Universal Robots URScript: FaiChun_9 Jan_11_2_t2.script

def Machining1():
  # Default parameters:
  global speed_ms = 0.05
  global speed_rads = 0.75
  global accel_mss = 3
  global accel_radss = 1.2
  global blend_radius_m = 0.0003

  # Add subprograms here
  # Start of main program
  # Program generated by RoboDK v5.6.8 for UR10e on 17/01/2025 16:04:48
  # Using nominal kinematics.
  blend_radius_m = 0.0003
  speed_ms = 0.05
  # set_reference(p[0.340000, -0.053000, 0.001500, 0.000000, 0.000000, 0.000000])
  set_tcp(p[0.000000, 0.000000, 0.252000, 0.000000, 0.000000, 0.000000])
  # Show Tool
  movej([0.537356, -1.385611, -2.455322, -0.871456, 1.570796, 2.108152],accel_radss,speed_rads,0,blend_radius_m)
  movel([0.537356, -1.438776, -2.485556, -0.788057, 1.570796, 2.108152],accel_mss,speed_ms,0,blend_radius_m)
  #SetTool1
  #M_RunCode6
  #SetRPM60000
  speed_ms = 0.05
  #M_RunCode3
  movel([0.537356, -1.461982, -2.496787, -0.753620, 1.570796, 2.108152],accel_mss,speed_ms,0,blend_radius_m)
  speed_ms = 0.003
  movel([0.537356, -1.467978, -2.499523, -0.744888, 1.570796, 2.108152],accel_mss,speed_ms,0,blend_radius_m)
  speed_ms = 0.02
  movel([0.264301, -1.461173, -2.505187, -0.746029, 1.570796, 1.835098],accel_mss,speed_ms,0,blend_radius_m)
  movel([0.376012, -1.125586, -2.705707, -0.881096, 1.570796, 1.946808],accel_mss,speed_ms,0,blend_radius_m)
  movel([0.747752, -1.141566, -2.699168, -0.871655, 1.570796, 2.318548],accel_mss,speed_ms,0,blend_radius_m)
  movel([0.537356, -1.467978, -2.499523, -0.744888, 1.570796, 2.108152],accel_mss,speed_ms,0,blend_radius_m)
  speed_ms = 0.003
  movel([0.537356, -1.461982, -2.496787, -0.753620, 1.570796, 2.108152],accel_mss,speed_ms,0,blend_radius_m)
  speed_ms = 0.05
  movel([0.537356, -1.438776, -2.485556, -0.788057, 1.570796, 2.108152],accel_mss,speed_ms,0,blend_radius_m)
  #M_RunCode9
  movel([0.537227, -1.429917, -2.492594, -0.789878, 1.570796, 2.108023],accel_mss,speed_ms,0,blend_radius_m)
  #M_RunCode3
  movel([0.537227, -1.453304, -2.503930, -0.755154, 1.570796, 2.108023],accel_mss,speed_ms,0,blend_radius_m)
  speed_ms = 0.003
  movel([0.537227, -1.459350, -2.506693, -0.746346, 1.570796, 2.108023],accel_mss,speed_ms,0,blend_radius_m)
  speed_ms = 0.012
  movel([0.533373, -1.458727, -2.507206, -0.746456, 1.570796, 2.104169],accel_mss,speed_ms,0,blend_radius_m)
  movel([0.531104, -1.462629, -2.503981, -0.745779, 1.570796, 2.101900],accel_mss,speed_ms,0,blend_radius_m)
  movel([0.525395, -1.461744, -2.504715, -0.745930, 1.570796, 2.096191],accel_mss,speed_ms,0,blend_radius_m)
  movel([0.527644, -1.457831, -2.507943, -0.746615, 1.570796, 2.098440],accel_mss,speed_ms,0,blend_radius_m)
  movel([0.525630, -1.457526, -2.508194, -0.746669, 1.570796, 2.096426],accel_mss,speed_ms,0,blend_radius_m)
  movel([0.523386, -1.461442, -2.504965, -0.745982, 1.570796, 2.094182],accel_mss,speed_ms,0,blend_radius_m)
  movel([0.518575, -1.460738, -2.505547, -0.746104, 1.570796, 2.089372],accel_mss,speed_ms,0,blend_radius_m)
  movel([0.517641, -1.460602, -2.505659, -0.746128, 1.570796, 2.088438],accel_mss,speed_ms,0,blend_radius_m)
  movel([0.520940, -1.454785, -2.510440, -0.747164, 1.570796, 2.091736],accel_mss,speed_ms,0,blend_radius_m)
  movel([0.524842, -1.455357, -2.509972, -0.747060, 1.570796, 2.095639],accel_mss,speed_ms,0,blend_radius_m)
  movel([0.526016, -1.453307, -2.511646, -0.747436, 1.570796, 2.096813],accel_mss,speed_ms,0,blend_radius_m)
  movel([0.520074, -1.452441, -2.512352, -0.747596, 1.570796, 2.090870],accel_mss,speed_ms,0,blend_radius_m)
  movel([0.515622, -1.460318, -2.505894, -0.746177, 1.570796, 2.086418],accel_mss,speed_ms,0,blend_radius_m)
  movel([0.514683, -1.460189, -2.506001, -0.746199, 1.570796, 2.085480],accel_mss,speed_ms,0,blend_radius_m)
  speed_ms = 0.02
  movel([0.406474, -1.451431, -2.513173, -0.747785, 1.570796, 1.977270],accel_mss,speed_ms,0,blend_radius_m)
  movel([0.291548, -1.454758, -2.510462, -0.747169, 1.570796, 1.862344],accel_mss,speed_ms,0,blend_radius_m)
  speed_ms = 0.012
  movel([0.294155, -1.446765, -2.516946, -0.748678, 1.570796, 1.864951],accel_mss,speed_ms,0,blend_radius_m)
  movel([0.287539, -1.447324, -2.516496, -0.748569, 1.570796, 1.858335],accel_mss,speed_ms,0,blend_radius_m)
  movel([0.286869, -1.449403, -2.514817, -0.748169, 1.570796, 1.857666],accel_mss,speed_ms,0,blend_radius_m)
  movel([0.291218, -1.449032, -2.515117, -0.748240, 1.570796, 1.862014],accel_mss,speed_ms,0,blend_radius_m)
  movel([0.289302, -1.454935, -2.510317, -0.747137, 1.570796, 1.860098],accel_mss,speed_ms,0,blend_radius_m)
  movel([0.288263, -1.455022, -2.510246, -0.747121, 1.570796, 1.859059],accel_mss,speed_ms,0,blend_radius_m)
  movel([0.282904, -1.455482, -2.509870, -0.747037, 1.570796, 1.853700],accel_mss,speed_ms,0,blend_radius_m)
  movel([0.284166, -1.451508, -2.513110, -0.747771, 1.570796, 1.854962],accel_mss,speed_ms,0,blend_radius_m)
  movel([0.281913, -1.451708, -2.512947, -0.747733, 1.570796, 1.852710],accel_mss,speed_ms,0,blend_radius_m)
  movel([0.280661, -1.455682, -2.509706, -0.747001, 1.570796, 1.851457],accel_mss,speed_ms,0,blend_radius_m)
  movel([0.274256, -1.456275, -2.509221, -0.746894, 1.570796, 1.845052],accel_mss,speed_ms,0,blend_radius_m)
  movel([0.275479, -1.452309, -2.512459, -0.747621, 1.570796, 1.846276],accel_mss,speed_ms,0,blend_radius_m)
  movel([0.271129, -1.452735, -2.512112, -0.747542, 1.570796, 1.841925],accel_mss,speed_ms,0,blend_radius_m)
  movel([0.272932, -1.446825, -2.516897, -0.748666, 1.570796, 1.843728],accel_mss,speed_ms,0,blend_radius_m)
  movel([0.277309, -1.446393, -2.517245, -0.748750, 1.570796, 1.848106],accel_mss,speed_ms,0,blend_radius_m)
  movel([0.277957, -1.444307, -2.518920, -0.749161, 1.570796, 1.848754],accel_mss,speed_ms,0,blend_radius_m)
  movel([0.273570, -1.444740, -2.518573, -0.749076, 1.570796, 1.844366],accel_mss,speed_ms,0,blend_radius_m)
  movel([0.275104, -1.439738, -2.522566, -0.750085, 1.570796, 1.845900],accel_mss,speed_ms,0,blend_radius_m)
  movel([0.275407, -1.438760, -2.523343, -0.750287, 1.570796, 1.846203],accel_mss,speed_ms,0,blend_radius_m)
  movel([0.281948, -1.438112, -2.523856, -0.750421, 1.570796, 1.852744],accel_mss,speed_ms,0,blend_radius_m)
  movel([0.280675, -1.442163, -2.520635, -0.749591, 1.570796, 1.851471],accel_mss,speed_ms,0,blend_radius_m)
  movel([0.282958, -1.441947, -2.520808, -0.749635, 1.570796, 1.853754],accel_mss,speed_ms,0,blend_radius_m)
  movel([0.284909, -1.435781, -2.525698, -0.750910, 1.570796, 1.855706],accel_mss,speed_ms,0,blend_radius_m)
  movel([0.276057, -1.436649, -2.525013, -0.750727, 1.570796, 1.846853],accel_mss,speed_ms,0,blend_radius_m)
  movel([0.315010, -1.315779, -2.609859, -0.786751, 1.570796, 1.885806],accel_mss,speed_ms,0,blend_radius_m)
  speed_ms = 0.02
  movel([0.366945, -1.166741, -2.688352, -0.857296, 1.570796, 1.937742],accel_mss,speed_ms,0,blend_radius_m)
  movel([0.367496, -1.165223, -2.689023, -0.858143, 1.570796, 1.938292],accel_mss,speed_ms,0,blend_radius_m)
  speed_ms = 0.012
  movel([0.379333, -1.163455, -2.689801, -0.859133, 1.570796, 1.950130],accel_mss,speed_ms,0,blend_radius_m)
  movel([0.382947, -1.153742, -2.694017, -0.864630, 1.570796, 1.953743],accel_mss,speed_ms,0,blend_radius_m)
  movel([0.379852, -1.154196, -2.693822, -0.864371, 1.570796, 1.950648],accel_mss,speed_ms,0,blend_radius_m)
  movel([0.377482, -1.160600, -2.691050, -0.860739, 1.570796, 1.948278],accel_mss,speed_ms,0,blend_radius_m)
  movel([0.368695, -1.161928, -2.690470, -0.859991, 1.570796, 1.939492],accel_mss,speed_ms,0,blend_radius_m)
  movel([0.369247, -1.160401, -2.691137, -0.860851, 1.570796, 1.940044],accel_mss,speed_ms,0,blend_radius_m)
  movel([0.372128, -1.152454, -2.694569, -0.865366, 1.570796, 1.942924],accel_mss,speed_ms,0,blend_radius_m)
  movel([0.378119, -1.151528, -2.694965, -0.865896, 1.570796, 1.948915],accel_mss,speed_ms,0,blend_radius_m)
  movel([0.379358, -1.148166, -2.696395, -0.867829, 1.570796, 1.950154],accel_mss,speed_ms,0,blend_radius_m)
  movel([0.373347, -1.149100, -2.695999, -0.867291, 1.570796, 1.944143],accel_mss,speed_ms,0,blend_radius_m)
  movel([0.376872, -1.139423, -2.700060, -0.872907, 1.570796, 1.947669],accel_mss,speed_ms,0,blend_radius_m)
  movel([0.382941, -1.138466, -2.700456, -0.873467, 1.570796, 1.953738],accel_mss,speed_ms,0,blend_radius_m)
  movel([0.385401, -1.131831, -2.703181, -0.877377, 1.570796, 1.956197],accel_mss,speed_ms,0,blend_radius_m)
  movel([0.394435, -1.130456, -2.703741, -0.878193, 1.570796, 1.965231],accel_mss,speed_ms,0,blend_radius_m)
  movel([0.391917, -1.137114, -2.701015, -0.874260, 1.570796, 1.962713],accel_mss,speed_ms,0,blend_radius_m)
  movel([0.395057, -1.136658, -2.701203, -0.874528, 1.570796, 1.965853],accel_mss,speed_ms,0,blend_radius_m)
  movel([0.397596, -1.129993, -2.703928, -0.878468, 1.570796, 1.968392],accel_mss,speed_ms,0,blend_radius_m)
  movel([0.406602, -1.128726, -2.704442, -0.879221, 1.570796, 1.977398],accel_mss,speed_ms,0,blend_radius_m)
  movel([0.402769, -1.138603, -2.700399, -0.873387, 1.570796, 1.973565],accel_mss,speed_ms,0,blend_radius_m)
  movel([0.396746, -1.139429, -2.700057, -0.872903, 1.570796, 1.967543],accel_mss,speed_ms,0,blend_radius_m)
  movel([0.395440, -1.142849, -2.698632, -0.870908, 1.570796, 1.966236],accel_mss,speed_ms,0,blend_radius_m)
  movel([0.404555, -1.141619, -2.699146, -0.871624, 1.570796, 1.975351],accel_mss,speed_ms,0,blend_radius_m)
  movel([0.409752, -1.128301, -2.704613, -0.879474, 1.570796, 1.980548],accel_mss,speed_ms,0,blend_radius_m)
  movel([0.568735, -1.120522, -2.707727, -0.884139, 1.570796, 2.139531],accel_mss,speed_ms,0,blend_radius_m)
  speed_ms = 0.02
  movel([0.712082, -1.141087, -2.699368, -0.871934, 1.570796, 2.282879],accel_mss,speed_ms,0,blend_radius_m)
  movel([0.703666, -1.154003, -2.693905, -0.864481, 1.570796, 2.274462],accel_mss,speed_ms,0,blend_radius_m)
  speed_ms = 0.012
  movel([0.711078, -1.155876, -2.693099, -0.863414, 1.570796, 2.281874],accel_mss,speed_ms,0,blend_radius_m)
  movel([0.713256, -1.152569, -2.694520, -0.865300, 1.570796, 2.284052],accel_mss,speed_ms,0,blend_radius_m)
  movel([0.708376, -1.151318, -2.695054, -0.866017, 1.570796, 2.279173],accel_mss,speed_ms,0,blend_radius_m)
  movel([0.714644, -1.141751, -2.699091, -0.871547, 1.570796, 2.285440],accel_mss,speed_ms,0,blend_radius_m)
  movel([0.715827, -1.142057, -2.698963, -0.871369, 1.570796, 2.286624],accel_mss,speed_ms,0,blend_radius_m)
  movel([0.721900, -1.143661, -2.698292, -0.870436, 1.570796, 2.292696],accel_mss,speed_ms,0,blend_radius_m)
  movel([0.717633, -1.150105, -2.695571, -0.866713, 1.570796, 2.288429],accel_mss,speed_ms,0,blend_radius_m)
  movel([0.720150, -1.150783, -2.695282, -0.866323, 1.570796, 2.290946],accel_mss,speed_ms,0,blend_radius_m)
  movel([0.724433, -1.144348, -2.698004, -0.870037, 1.570796, 2.295229],accel_mss,speed_ms,0,blend_radius_m)
  movel([0.731605, -1.146355, -2.697160, -0.868874, 1.570796, 2.302401],accel_mss,speed_ms,0,blend_radius_m)
  movel([0.727300, -1.152759, -2.694438, -0.865192, 1.570796, 2.298096],accel_mss,speed_ms,0,blend_radius_m)
  movel([0.732091, -1.154132, -2.693850, -0.864408, 1.570796, 2.302888],accel_mss,speed_ms,0,blend_radius_m)
  movel([0.725789, -1.163458, -2.689799, -0.859132, 1.570796, 2.296585],accel_mss,speed_ms,0,blend_radius_m)
  movel([0.721022, -1.162117, -2.690387, -0.859885, 1.570796, 2.291818],accel_mss,speed_ms,0,blend_radius_m)
  movel([0.718847, -1.165363, -2.688961, -0.858065, 1.570796, 2.289644],accel_mss,speed_ms,0,blend_radius_m)
  movel([0.723604, -1.166697, -2.688372, -0.857320, 1.570796, 2.294400],accel_mss,speed_ms,0,blend_radius_m)
  movel([0.718442, -1.174360, -2.684951, -0.853078, 1.570796, 2.289239],accel_mss,speed_ms,0,blend_radius_m)
  movel([0.717449, -1.175836, -2.684285, -0.852268, 1.570796, 2.288246],accel_mss,speed_ms,0,blend_radius_m)
  movel([0.710428, -1.173922, -2.685148, -0.853319, 1.570796, 2.281224],accel_mss,speed_ms,0,blend_radius_m)
  movel([0.714548, -1.167736, -2.687912, -0.856742, 1.570796, 2.285344],accel_mss,speed_ms,0,blend_radius_m)
  movel([0.712062, -1.167070, -2.688207, -0.857112, 1.570796, 2.282858],accel_mss,speed_ms,0,blend_radius_m)
  movel([0.705834, -1.176462, -2.684002, -0.851925, 1.570796, 2.276630],accel_mss,speed_ms,0,blend_radius_m)
  movel([0.715315, -1.179011, -2.682845, -0.850533, 1.570796, 2.286112],accel_mss,speed_ms,0,blend_radius_m)
  speed_ms = 0.02
  movel([0.619516, -1.325160, -2.604003, -0.783226, 1.570796, 2.190312],accel_mss,speed_ms,0,blend_radius_m)
  movel([0.546569, -1.443533, -2.519541, -0.749316, 1.570796, 2.117365],accel_mss,speed_ms,0,blend_radius_m)
  speed_ms = 0.012
  movel([0.538730, -1.442256, -2.520561, -0.749572, 1.570796, 2.109526],accel_mss,speed_ms,0,blend_radius_m)
  movel([0.535189, -1.448324, -2.515689, -0.748376, 1.570796, 2.105985],accel_mss,speed_ms,0,blend_radius_m)
  movel([0.537216, -1.448646, -2.515429, -0.748314, 1.570796, 2.108012],accel_mss,speed_ms,0,blend_radius_m)
  movel([0.539548, -1.444662, -2.518636, -0.749091, 1.570796, 2.110344],accel_mss,speed_ms,0,blend_radius_m)
  movel([0.545329, -1.445610, -2.517875, -0.748904, 1.570796, 2.116125],accel_mss,speed_ms,0,blend_radius_m)
  movel([0.544761, -1.446568, -2.517104, -0.748716, 1.570796, 2.115557],accel_mss,speed_ms,0,blend_radius_m)
  movel([0.541852, -1.451489, -2.513125, -0.747774, 1.570796, 2.112648],accel_mss,speed_ms,0,blend_radius_m)
  movel([0.537972, -1.450854, -2.513641, -0.747894, 1.570796, 2.108768],accel_mss,speed_ms,0,blend_radius_m)
  movel([0.536771, -1.452905, -2.511974, -0.747510, 1.570796, 2.107567],accel_mss,speed_ms,0,blend_radius_m)
  movel([0.540646, -1.453538, -2.511458, -0.747393, 1.570796, 2.111442],accel_mss,speed_ms,0,blend_radius_m)
  movel([0.537227, -1.459350, -2.506693, -0.746346, 1.570796, 2.108023],accel_mss,speed_ms,0,blend_radius_m)
  speed_ms = 0.003
  movel([0.537227, -1.453304, -2.503930, -0.755154, 1.570796, 2.108023],accel_mss,speed_ms,0,blend_radius_m)
  speed_ms = 0.05
  movel([0.537227, -1.429917, -2.492594, -0.789878, 1.570796, 2.108023],accel_mss,speed_ms,0,blend_radius_m)
  #M_RunCode9
  movel([0.423144, -1.170555, -2.652350, -0.889483, 1.570796, 1.993941],accel_mss,speed_ms,0,blend_radius_m)
  #M_RunCode3
  # num 0 inside
  movel([0.423144, -1.197858, -2.667024, -0.847507, 1.570796, 1.993941],accel_mss,speed_ms,0,blend_radius_m)
  speed_ms = 0.003
  movel([0.423144, -1.205044, -2.670628, -0.836717, 1.570796, 1.993941],accel_mss,speed_ms,0,blend_radius_m)
  speed_ms = 0.015
  movel([0.414451, -1.211707, -2.667382, -0.833300, 1.570796, 1.985247],accel_mss,speed_ms,0,blend_radius_m)
  movel([0.408145, -1.215978, -2.665275, -0.831136, 1.570796, 1.978941],accel_mss,speed_ms,0,blend_radius_m)
  movel([0.405824, -1.217205, -2.664666, -0.830518, 1.570796, 1.976621],accel_mss,speed_ms,0,blend_radius_m)
  movel([0.403998, -1.217788, -2.664376, -0.830225, 1.570796, 1.974795],accel_mss,speed_ms,0,blend_radius_m)
  movel([0.402664, -1.217733, -2.664403, -0.830253, 1.570796, 1.973460],accel_mss,speed_ms,0,blend_radius_m)
  movel([0.401818, -1.217039, -2.664748, -0.830602, 1.570796, 1.972614],accel_mss,speed_ms,0,blend_radius_m)
  movel([0.401559, -1.215868, -2.665329, -0.831191, 1.570796, 1.972356],accel_mss,speed_ms,0,blend_radius_m)
  movel([0.401991, -1.214387, -2.666062, -0.831940, 1.570796, 1.972787],accel_mss,speed_ms,0,blend_radius_m)
  movel([0.403116, -1.212593, -2.666947, -0.832850, 1.570796, 1.973912],accel_mss,speed_ms,0,blend_radius_m)
  movel([0.404937, -1.210479, -2.667984, -0.833926, 1.570796, 1.975733],accel_mss,speed_ms,0,blend_radius_m)
  movel([0.410670, -1.205076, -2.670613, -0.836701, 1.570796, 1.981466],accel_mss,speed_ms,0,blend_radius_m)
  movel([0.419217, -1.197936, -2.674037, -0.840416, 1.570796, 1.990013],accel_mss,speed_ms,0,blend_radius_m)
  movel([0.428065, -1.191105, -2.677261, -0.844024, 1.570796, 1.998861],accel_mss,speed_ms,0,blend_radius_m)
  movel([0.434586, -1.186692, -2.679317, -0.846381, 1.570796, 2.005382],accel_mss,speed_ms,0,blend_radius_m)
  movel([0.436993, -1.185433, -2.679899, -0.847057, 1.570796, 2.007789],accel_mss,speed_ms,0,blend_radius_m)
  movel([0.438876, -1.184846, -2.680170, -0.847373, 1.570796, 2.009672],accel_mss,speed_ms,0,blend_radius_m)
  movel([0.440232, -1.184936, -2.680129, -0.847325, 1.570796, 2.011028],accel_mss,speed_ms,0,blend_radius_m)
  movel([0.441059, -1.185700, -2.679775, -0.846913, 1.570796, 2.011856],accel_mss,speed_ms,0,blend_radius_m)
  movel([0.441266, -1.186954, -2.679195, -0.846240, 1.570796, 2.012062],accel_mss,speed_ms,0,blend_radius_m)
  movel([0.440764, -1.188513, -2.678471, -0.845406, 1.570796, 2.011560],accel_mss,speed_ms,0,blend_radius_m)
  movel([0.439549, -1.190375, -2.677602, -0.844412, 1.570796, 2.010346],accel_mss,speed_ms,0,blend_radius_m)
  movel([0.437636, -1.192534, -2.676590, -0.843265, 1.570796, 2.008432],accel_mss,speed_ms,0,blend_radius_m)
  movel([0.431736, -1.197976, -2.674018, -0.840395, 1.570796, 2.002532],accel_mss,speed_ms,0,blend_radius_m)
  movel([0.423144, -1.205044, -2.670628, -0.836717, 1.570796, 1.993941],accel_mss,speed_ms,0,blend_radius_m)
  speed_ms = 0.003
  movel([0.423144, -1.197858, -2.667024, -0.847507, 1.570796, 1.993941],accel_mss,speed_ms,0,blend_radius_m)
  speed_ms = 0.05
  movel([0.423144, -1.170555, -2.652350, -0.889483, 1.570796, 1.993941],accel_mss,speed_ms,0,blend_radius_m)
  #M_RunCode9
  movel([0.427307, -1.178294, -2.648743, -0.885352, 1.570796, 1.998103],accel_mss,speed_ms,0,blend_radius_m)
  #M_RunCode3
  #num 0 outside
  movel([0.427307, -1.205537, -2.663314, -0.843537, 1.570796, 1.998103],accel_mss,speed_ms,0,blend_radius_m)
  speed_ms = 0.003
  movel([0.427307, -1.212702, -2.666893, -0.832794, 1.570796, 1.998103],accel_mss,speed_ms,0,blend_radius_m)
  speed_ms = 0.015
  movel([0.424140, -1.215057, -2.665731, -0.831601, 1.570796, 1.994936],accel_mss,speed_ms,0,blend_radius_m)
  movel([0.421112, -1.217044, -2.664746, -0.830599, 1.570796, 1.991909],accel_mss,speed_ms,0,blend_radius_m)
  movel([0.418216, -1.218671, -2.663936, -0.829782, 1.570796, 1.989013],accel_mss,speed_ms,0,blend_radius_m)
  movel([0.415452, -1.219937, -2.663303, -0.829148, 1.570796, 1.986248],accel_mss,speed_ms,0,blend_radius_m)
  movel([0.412856, -1.220852, -2.662845, -0.828692, 1.570796, 1.983652],accel_mss,speed_ms,0,blend_radius_m)
  movel([0.410467, -1.221421, -2.662560, -0.828408, 1.570796, 1.981263],accel_mss,speed_ms,0,blend_radius_m)
  movel([0.408281, -1.221649, -2.662445, -0.828295, 1.570796, 1.979077],accel_mss,speed_ms,0,blend_radius_m)
  movel([0.406301, -1.221529, -2.662506, -0.828354, 1.570796, 1.977097],accel_mss,speed_ms,0,blend_radius_m)
  movel([0.404543, -1.221083, -2.662730, -0.828577, 1.570796, 1.975339],accel_mss,speed_ms,0,blend_radius_m)
  movel([0.403031, -1.220334, -2.663105, -0.828950, 1.570796, 1.973827],accel_mss,speed_ms,0,blend_radius_m)
  movel([0.401762, -1.219277, -2.663633, -0.829479, 1.570796, 1.972558],accel_mss,speed_ms,0,blend_radius_m)
  movel([0.400735, -1.217914, -2.664313, -0.830162, 1.570796, 1.971531],accel_mss,speed_ms,0,blend_radius_m)
  movel([0.399997, -1.216311, -2.665110, -0.830968, 1.570796, 1.970793],accel_mss,speed_ms,0,blend_radius_m)
  movel([0.399595, -1.214545, -2.665984, -0.831860, 1.570796, 1.970391],accel_mss,speed_ms,0,blend_radius_m)
  movel([0.399526, -1.212615, -2.666936, -0.832838, 1.570796, 1.970323],accel_mss,speed_ms,0,blend_radius_m)
  movel([0.399800, -1.210512, -2.667968, -0.833909, 1.570796, 1.970597],accel_mss,speed_ms,0,blend_radius_m)
  movel([0.400424, -1.208271, -2.669062, -0.835056, 1.570796, 1.971220],accel_mss,speed_ms,0,blend_radius_m)
  movel([0.401410, -1.205920, -2.670204, -0.836265, 1.570796, 1.972206],accel_mss,speed_ms,0,blend_radius_m)
  movel([0.402761, -1.203455, -2.671395, -0.837539, 1.570796, 1.973557],accel_mss,speed_ms,0,blend_radius_m)
  movel([0.404482, -1.200878, -2.672633, -0.838879, 1.570796, 1.975278],accel_mss,speed_ms,0,blend_radius_m)
  movel([0.406561, -1.198233, -2.673896, -0.840261, 1.570796, 1.977357],accel_mss,speed_ms,0,blend_radius_m)
  movel([0.408989, -1.195574, -2.675157, -0.841658, 1.570796, 1.979785],accel_mss,speed_ms,0,blend_radius_m)
  movel([0.411765, -1.192904, -2.676417, -0.843069, 1.570796, 1.982561],accel_mss,speed_ms,0,blend_radius_m)
  movel([0.414891, -1.190223, -2.677673, -0.844493, 1.570796, 1.985687],accel_mss,speed_ms,0,blend_radius_m)
  movel([0.418140, -1.187719, -2.678840, -0.845830, 1.570796, 1.988936],accel_mss,speed_ms,0,blend_radius_m)
  movel([0.421270, -1.185591, -2.679826, -0.846972, 1.570796, 1.992066],accel_mss,speed_ms,0,blend_radius_m)
  movel([0.424280, -1.183839, -2.680634, -0.847915, 1.570796, 1.995076],accel_mss,speed_ms,0,blend_radius_m)
  movel([0.427162, -1.182472, -2.681263, -0.848654, 1.570796, 1.997958],accel_mss,speed_ms,0,blend_radius_m)
  movel([0.429870, -1.181487, -2.681714, -0.849188, 1.570796, 2.000666],accel_mss,speed_ms,0,blend_radius_m)
  movel([0.432350, -1.180886, -2.681989, -0.849514, 1.570796, 2.003146],accel_mss,speed_ms,0,blend_radius_m)
  movel([0.434606, -1.180663, -2.682091, -0.849635, 1.570796, 2.005402],accel_mss,speed_ms,0,blend_radius_m)
  movel([0.436631, -1.180826, -2.682017, -0.849547, 1.570796, 2.007428],accel_mss,speed_ms,0,blend_radius_m)
  movel([0.438404, -1.181343, -2.681780, -0.849266, 1.570796, 2.009201],accel_mss,speed_ms,0,blend_radius_m)
  movel([0.439913, -1.182188, -2.681393, -0.848808, 1.570796, 2.010710],accel_mss,speed_ms,0,blend_radius_m)
  movel([0.441158, -1.183359, -2.680855, -0.848175, 1.570796, 2.011954],accel_mss,speed_ms,0,blend_radius_m)
  movel([0.442132, -1.184852, -2.680167, -0.847370, 1.570796, 2.012929],accel_mss,speed_ms,0,blend_radius_m)
  movel([0.442800, -1.186585, -2.679366, -0.846438, 1.570796, 2.013596],accel_mss,speed_ms,0,blend_radius_m)
  movel([0.443122, -1.188471, -2.678490, -0.845428, 1.570796, 2.013919],accel_mss,speed_ms,0,blend_radius_m)
  movel([0.443100, -1.190509, -2.677539, -0.844340, 1.570796, 2.013897],accel_mss,speed_ms,0,blend_radius_m)
  movel([0.442736, -1.192698, -2.676513, -0.843178, 1.570796, 2.013532],accel_mss,speed_ms,0,blend_radius_m)
  movel([0.442021, -1.195002, -2.675428, -0.841959, 1.570796, 2.012817],accel_mss,speed_ms,0,blend_radius_m)
  movel([0.440945, -1.197394, -2.674295, -0.840701, 1.570796, 2.011742],accel_mss,speed_ms,0,blend_radius_m)
  movel([0.439509, -1.199872, -2.673114, -0.839403, 1.570796, 2.010305],accel_mss,speed_ms,0,blend_radius_m)
  movel([0.437718, -1.202433, -2.671886, -0.838069, 1.570796, 2.008514],accel_mss,speed_ms,0,blend_radius_m)
  movel([0.435592, -1.205026, -2.670637, -0.836727, 1.570796, 2.006388],accel_mss,speed_ms,0,blend_radius_m)
  movel([0.433145, -1.207602, -2.669388, -0.835400, 1.570796, 2.003941],accel_mss,speed_ms,0,blend_radius_m)
  movel([0.430383, -1.210160, -2.668140, -0.834089, 1.570796, 2.001179],accel_mss,speed_ms,0,blend_radius_m)
  movel([0.427307, -1.212702, -2.666893, -0.832794, 1.570796, 1.998103],accel_mss,speed_ms,0,blend_radius_m)
  speed_ms = 0.003
  movel([0.427307, -1.205537, -2.663314, -0.843537, 1.570796, 1.998103],accel_mss,speed_ms,0,blend_radius_m)
  speed_ms = 0.05
  movel([0.427307, -1.178294, -2.648743, -0.885352, 1.570796, 1.998103],accel_mss,speed_ms,0,blend_radius_m)
  #M_RunCode9
  movel([0.404280, -1.160081, -2.657135, -0.895174, 1.570796, 1.975076],accel_mss,speed_ms,0,blend_radius_m)
  #M_RunCode3
  movel([0.404280, -1.187457, -2.671946, -0.852986, 1.570796, 1.975076],accel_mss,speed_ms,0,blend_radius_m)
  speed_ms = 0.003
  movel([0.404280, -1.194669, -2.675585, -0.842135, 1.570796, 1.975076],accel_mss,speed_ms,0,blend_radius_m)
  speed_ms = 0.02
  movel([0.393218, -1.203772, -2.671242, -0.837375, 1.570796, 1.964014],accel_mss,speed_ms,0,blend_radius_m)
  movel([0.379156, -1.181402, -2.681753, -0.849234, 1.570796, 1.949952],accel_mss,speed_ms,0,blend_radius_m)
  movel([0.380274, -1.180444, -2.682191, -0.849754, 1.570796, 1.951070],accel_mss,speed_ms,0,blend_radius_m)
  movel([0.383293, -1.178260, -2.683187, -0.850943, 1.570796, 1.954090],accel_mss,speed_ms,0,blend_radius_m)
  movel([0.386594, -1.176640, -2.683921, -0.851828, 1.570796, 1.957391],accel_mss,speed_ms,0,blend_radius_m)
  movel([0.390000, -1.175505, -2.684435, -0.852450, 1.570796, 1.960797],accel_mss,speed_ms,0,blend_radius_m)
  movel([0.393328, -1.174770, -2.684766, -0.852853, 1.570796, 1.964124],accel_mss,speed_ms,0,blend_radius_m)
  movel([0.401978, -1.173719, -2.685239, -0.853430, 1.570796, 1.972774],accel_mss,speed_ms,0,blend_radius_m)
  movel([0.409948, -1.172895, -2.685609, -0.853884, 1.570796, 1.980745],accel_mss,speed_ms,0,blend_radius_m)
  movel([0.413040, -1.172290, -2.685881, -0.854218, 1.570796, 1.983837],accel_mss,speed_ms,0,blend_radius_m)
  movel([0.416142, -1.171341, -2.686306, -0.854742, 1.570796, 1.986939],accel_mss,speed_ms,0,blend_radius_m)
  movel([0.419104, -1.169981, -2.686913, -0.855494, 1.570796, 1.989900],accel_mss,speed_ms,0,blend_radius_m)
  movel([0.421778, -1.168142, -2.687732, -0.856516, 1.570796, 1.992574],accel_mss,speed_ms,0,blend_radius_m)
  movel([0.424597, -1.165348, -2.688967, -0.858073, 1.570796, 1.995393],accel_mss,speed_ms,0,blend_radius_m)
  movel([0.425571, -1.163955, -2.689581, -0.858853, 1.570796, 1.996367],accel_mss,speed_ms,0,blend_radius_m)
  movel([0.426254, -1.162565, -2.690191, -0.859633, 1.570796, 1.997050],accel_mss,speed_ms,0,blend_radius_m)
  movel([0.426823, -1.160031, -2.691298, -0.861060, 1.570796, 1.997619],accel_mss,speed_ms,0,blend_radius_m)
  movel([0.426371, -1.158003, -2.692179, -0.862207, 1.570796, 1.997167],accel_mss,speed_ms,0,blend_radius_m)
  movel([0.425588, -1.157027, -2.692602, -0.862760, 1.570796, 1.996384],accel_mss,speed_ms,0,blend_radius_m)
  movel([0.424615, -1.156628, -2.692774, -0.862986, 1.570796, 1.995411],accel_mss,speed_ms,0,blend_radius_m)
  movel([0.423553, -1.156764, -2.692715, -0.862910, 1.570796, 1.994350],accel_mss,speed_ms,0,blend_radius_m)
  movel([0.422516, -1.157377, -2.692450, -0.862562, 1.570796, 1.993312],accel_mss,speed_ms,0,blend_radius_m)
  movel([0.421350, -1.158935, -2.691775, -0.861679, 1.570796, 1.992147],accel_mss,speed_ms,0,blend_radius_m)
  movel([0.420302, -1.160502, -2.691093, -0.860794, 1.570796, 1.991098],accel_mss,speed_ms,0,blend_radius_m)
  movel([0.418652, -1.162130, -2.690381, -0.859877, 1.570796, 1.989448],accel_mss,speed_ms,0,blend_radius_m)
  movel([0.416433, -1.163562, -2.689754, -0.859074, 1.570796, 1.987229],accel_mss,speed_ms,0,blend_radius_m)
  movel([0.414428, -1.164000, -2.689561, -0.858828, 1.570796, 1.985224],accel_mss,speed_ms,0,blend_radius_m)
  movel([0.412782, -1.163572, -2.689749, -0.859068, 1.570796, 1.983579],accel_mss,speed_ms,0,blend_radius_m)
  movel([0.411645, -1.162404, -2.690262, -0.859724, 1.570796, 1.982442],accel_mss,speed_ms,0,blend_radius_m)
  movel([0.411141, -1.160707, -2.691003, -0.860679, 1.570796, 1.981937],accel_mss,speed_ms,0,blend_radius_m)
  movel([0.411392, -1.158682, -2.691885, -0.861822, 1.570796, 1.982188],accel_mss,speed_ms,0,blend_radius_m)
  movel([0.412449, -1.156544, -2.692811, -0.863035, 1.570796, 1.983246],accel_mss,speed_ms,0,blend_radius_m)
  movel([0.414364, -1.154517, -2.693684, -0.864188, 1.570796, 1.985161],accel_mss,speed_ms,0,blend_radius_m)
  movel([0.416288, -1.153142, -2.694274, -0.864973, 1.570796, 1.987084],accel_mss,speed_ms,0,blend_radius_m)
  movel([0.418172, -1.152282, -2.694642, -0.865464, 1.570796, 1.988968],accel_mss,speed_ms,0,blend_radius_m)
  movel([0.420018, -1.151940, -2.694789, -0.865661, 1.570796, 1.990814],accel_mss,speed_ms,0,blend_radius_m)
  movel([0.421820, -1.152122, -2.694711, -0.865556, 1.570796, 1.992616],accel_mss,speed_ms,0,blend_radius_m)
  movel([0.423510, -1.152764, -2.694436, -0.865189, 1.570796, 1.994306],accel_mss,speed_ms,0,blend_radius_m)
  movel([0.425030, -1.153795, -2.693994, -0.864600, 1.570796, 1.995826],accel_mss,speed_ms,0,blend_radius_m)
  movel([0.427544, -1.157036, -2.692598, -0.862755, 1.570796, 1.998341],accel_mss,speed_ms,0,blend_radius_m)
  movel([0.428643, -1.159554, -2.691506, -0.861329, 1.570796, 1.999440],accel_mss,speed_ms,0,blend_radius_m)
  movel([0.429311, -1.162232, -2.690337, -0.859820, 1.570796, 2.000108],accel_mss,speed_ms,0,blend_radius_m)
  movel([0.429551, -1.165062, -2.689094, -0.858233, 1.570796, 2.000347],accel_mss,speed_ms,0,blend_radius_m)
  movel([0.429364, -1.168043, -2.687775, -0.856571, 1.570796, 2.000160],accel_mss,speed_ms,0,blend_radius_m)
  movel([0.428602, -1.171050, -2.686436, -0.854903, 1.570796, 1.999398],accel_mss,speed_ms,0,blend_radius_m)
  movel([0.427100, -1.173969, -2.685127, -0.853293, 1.570796, 1.997897],accel_mss,speed_ms,0,blend_radius_m)
  movel([0.424869, -1.176799, -2.683850, -0.851741, 1.570796, 1.995665],accel_mss,speed_ms,0,blend_radius_m)
  movel([0.421913, -1.179542, -2.682603, -0.850244, 1.570796, 1.992710],accel_mss,speed_ms,0,blend_radius_m)
  movel([0.418973, -1.181635, -2.681646, -0.849107, 1.570796, 1.989769],accel_mss,speed_ms,0,blend_radius_m)
  movel([0.416007, -1.183151, -2.680951, -0.848287, 1.570796, 1.986803],accel_mss,speed_ms,0,blend_radius_m)
  movel([0.413084, -1.184191, -2.680472, -0.847726, 1.570796, 1.983881],accel_mss,speed_ms,0,blend_radius_m)
  movel([0.410281, -1.184855, -2.680166, -0.847368, 1.570796, 1.981077],accel_mss,speed_ms,0,blend_radius_m)
  movel([0.403638, -1.185636, -2.679805, -0.846948, 1.570796, 1.974434],accel_mss,speed_ms,0,blend_radius_m)
  movel([0.397343, -1.186447, -2.679430, -0.846512, 1.570796, 1.968140],accel_mss,speed_ms,0,blend_radius_m)
  movel([0.394791, -1.187071, -2.679141, -0.846178, 1.570796, 1.965587],accel_mss,speed_ms,0,blend_radius_m)
  movel([0.392175, -1.188020, -2.678700, -0.845669, 1.570796, 1.962972],accel_mss,speed_ms,0,blend_radius_m)
  movel([0.389578, -1.189370, -2.678071, -0.844948, 1.570796, 1.960374],accel_mss,speed_ms,0,blend_radius_m)
  movel([0.387093, -1.191182, -2.677224, -0.843982, 1.570796, 1.957889],accel_mss,speed_ms,0,blend_radius_m)
  movel([0.387619, -1.192022, -2.676831, -0.843536, 1.570796, 1.958415],accel_mss,speed_ms,0,blend_radius_m)
  movel([0.389239, -1.194207, -2.675803, -0.842379, 1.570796, 1.960035],accel_mss,speed_ms,0,blend_radius_m)
  movel([0.391018, -1.195821, -2.675040, -0.841528, 1.570796, 1.961815],accel_mss,speed_ms,0,blend_radius_m)
  movel([0.392953, -1.196869, -2.674543, -0.840976, 1.570796, 1.963749],accel_mss,speed_ms,0,blend_radius_m)
  movel([0.395052, -1.197352, -2.674314, -0.840723, 1.570796, 1.965848],accel_mss,speed_ms,0,blend_radius_m)
  movel([0.397259, -1.197336, -2.674322, -0.840731, 1.570796, 1.968056],accel_mss,speed_ms,0,blend_radius_m)
  movel([0.399531, -1.196885, -2.674536, -0.840968, 1.570796, 1.970328],accel_mss,speed_ms,0,blend_radius_m)
  movel([0.401868, -1.195997, -2.674957, -0.841435, 1.570796, 1.972665],accel_mss,speed_ms,0,blend_radius_m)
  movel([0.404280, -1.194669, -2.675585, -0.842135, 1.570796, 1.975076],accel_mss,speed_ms,0,blend_radius_m)
  speed_ms = 0.003
  movel([0.404280, -1.187457, -2.671946, -0.852986, 1.570796, 1.975076],accel_mss,speed_ms,0,blend_radius_m)
  speed_ms = 0.05
  movel([0.404280, -1.160081, -2.657135, -0.895174, 1.570796, 1.975076],accel_mss,speed_ms,0,blend_radius_m)
  #M_RunCode9
  movel([0.496458, -1.374956, -2.533748, -0.803685, 1.570796, 2.067255],accel_mss,speed_ms,0,blend_radius_m)
  #M_RunCode3
  movel([0.496458, -1.399421, -2.545759, -0.767209, 1.570796, 2.067255],accel_mss,speed_ms,0,blend_radius_m)
  speed_ms = 0.003
  movel([0.496458, -1.405765, -2.548690, -0.757933, 1.570796, 2.067255],accel_mss,speed_ms,0,blend_radius_m)
  speed_ms = 0.02
  movel([0.498829, -1.404633, -2.549531, -0.758224, 1.570796, 2.069626],accel_mss,speed_ms,0,blend_radius_m)
  movel([0.501342, -1.403976, -2.550019, -0.758394, 1.570796, 2.072138],accel_mss,speed_ms,0,blend_radius_m)
  movel([0.503880, -1.403701, -2.550223, -0.758465, 1.570796, 2.074676],accel_mss,speed_ms,0,blend_radius_m)
  movel([0.506317, -1.403718, -2.550210, -0.758461, 1.570796, 2.077114],accel_mss,speed_ms,0,blend_radius_m)
  movel([0.512569, -1.404395, -2.549708, -0.758286, 1.570796, 2.083365],accel_mss,speed_ms,0,blend_radius_m)
  movel([0.518313, -1.405116, -2.549173, -0.758100, 1.570796, 2.089109],accel_mss,speed_ms,0,blend_radius_m)
  movel([0.520565, -1.405182, -2.549124, -0.758083, 1.570796, 2.091362],accel_mss,speed_ms,0,blend_radius_m)
  movel([0.522857, -1.404990, -2.549267, -0.758132, 1.570796, 2.093653],accel_mss,speed_ms,0,blend_radius_m)
  movel([0.525085, -1.404469, -2.549653, -0.758267, 1.570796, 2.095881],accel_mss,speed_ms,0,blend_radius_m)
  movel([0.527150, -1.403543, -2.550339, -0.758506, 1.570796, 2.097946],accel_mss,speed_ms,0,blend_radius_m)
  movel([0.529402, -1.401935, -2.551529, -0.758926, 1.570796, 2.100198],accel_mss,speed_ms,0,blend_radius_m)
  movel([0.530218, -1.401063, -2.552172, -0.759155, 1.570796, 2.101014],accel_mss,speed_ms,0,blend_radius_m)
  movel([0.530826, -1.400145, -2.552847, -0.759397, 1.570796, 2.101623],accel_mss,speed_ms,0,blend_radius_m)
  movel([0.531457, -1.398361, -2.554157, -0.759871, 1.570796, 2.102253],accel_mss,speed_ms,0,blend_radius_m)
  movel([0.531320, -1.396783, -2.555312, -0.760294, 1.570796, 2.102116],accel_mss,speed_ms,0,blend_radius_m)
  movel([0.530856, -1.395926, -2.555937, -0.760525, 1.570796, 2.101653],accel_mss,speed_ms,0,blend_radius_m)
  movel([0.530202, -1.395470, -2.556270, -0.760649, 1.570796, 2.100998],accel_mss,speed_ms,0,blend_radius_m)
  movel([0.529443, -1.395389, -2.556329, -0.760671, 1.570796, 2.100239],accel_mss,speed_ms,0,blend_radius_m)
  movel([0.528654, -1.395669, -2.556125, -0.760595, 1.570796, 2.099451],accel_mss,speed_ms,0,blend_radius_m)
  movel([0.527688, -1.396628, -2.555425, -0.760336, 1.570796, 2.098485],accel_mss,speed_ms,0,blend_radius_m)
  movel([0.526802, -1.397617, -2.554702, -0.760070, 1.570796, 2.097599],accel_mss,speed_ms,0,blend_radius_m)
  movel([0.525485, -1.398548, -2.554020, -0.759821, 1.570796, 2.096281],accel_mss,speed_ms,0,blend_radius_m)
  movel([0.523783, -1.399242, -2.553511, -0.759636, 1.570796, 2.094579],accel_mss,speed_ms,0,blend_radius_m)
  movel([0.522323, -1.399228, -2.553521, -0.759640, 1.570796, 2.093120],accel_mss,speed_ms,0,blend_radius_m)
  movel([0.521196, -1.398631, -2.553959, -0.759799, 1.570796, 2.091992],accel_mss,speed_ms,0,blend_radius_m)
  movel([0.520501, -1.397571, -2.554736, -0.760082, 1.570796, 2.091298],accel_mss,speed_ms,0,blend_radius_m)
  movel([0.520305, -1.396218, -2.555724, -0.760446, 1.570796, 2.091102],accel_mss,speed_ms,0,blend_radius_m)
  movel([0.520673, -1.394753, -2.556792, -0.760844, 1.570796, 2.091470],accel_mss,speed_ms,0,blend_radius_m)
  movel([0.521620, -1.393344, -2.557816, -0.761229, 1.570796, 2.092417],accel_mss,speed_ms,0,blend_radius_m)
  movel([0.523162, -1.392165, -2.558670, -0.761553, 1.570796, 2.093958],accel_mss,speed_ms,0,blend_radius_m)
  movel([0.524646, -1.391470, -2.559173, -0.761746, 1.570796, 2.095442],accel_mss,speed_ms,0,blend_radius_m)
  movel([0.526056, -1.391155, -2.559401, -0.761833, 1.570796, 2.096853],accel_mss,speed_ms,0,blend_radius_m)
  movel([0.527388, -1.391218, -2.559355, -0.761816, 1.570796, 2.098184],accel_mss,speed_ms,0,blend_radius_m)
  movel([0.528640, -1.391659, -2.559037, -0.761693, 1.570796, 2.099436],accel_mss,speed_ms,0,blend_radius_m)
  movel([0.529774, -1.392419, -2.558487, -0.761484, 1.570796, 2.100570],accel_mss,speed_ms,0,blend_radius_m)
  movel([0.530751, -1.393442, -2.557745, -0.761202, 1.570796, 2.101547],accel_mss,speed_ms,0,blend_radius_m)
  movel([0.532237, -1.396261, -2.555693, -0.760435, 1.570796, 2.103034],accel_mss,speed_ms,0,blend_radius_m)
  movel([0.532787, -1.398311, -2.554194, -0.759884, 1.570796, 2.103583],accel_mss,speed_ms,0,blend_radius_m)
  movel([0.533020, -1.400406, -2.552656, -0.759328, 1.570796, 2.103817],accel_mss,speed_ms,0,blend_radius_m)
  movel([0.532938, -1.402543, -2.551079, -0.758767, 1.570796, 2.103734],accel_mss,speed_ms,0,blend_radius_m)
  movel([0.532540, -1.404724, -2.549464, -0.758201, 1.570796, 2.103336],accel_mss,speed_ms,0,blend_radius_m)
  movel([0.531729, -1.406831, -2.547897, -0.757661, 1.570796, 2.102526],accel_mss,speed_ms,0,blend_radius_m)
  movel([0.530402, -1.408755, -2.546460, -0.757174, 1.570796, 2.101198],accel_mss,speed_ms,0,blend_radius_m)
  movel([0.528563, -1.410498, -2.545154, -0.756737, 1.570796, 2.099359],accel_mss,speed_ms,0,blend_radius_m)
  movel([0.526209, -1.412062, -2.543978, -0.756349, 1.570796, 2.097006],accel_mss,speed_ms,0,blend_radius_m)
  movel([0.523926, -1.413146, -2.543161, -0.756082, 1.570796, 2.094722],accel_mss,speed_ms,0,blend_radius_m)
  movel([0.521671, -1.413796, -2.542670, -0.755923, 1.570796, 2.092468],accel_mss,speed_ms,0,blend_radius_m)
  movel([0.519488, -1.414096, -2.542444, -0.755850, 1.570796, 2.090284],accel_mss,speed_ms,0,blend_radius_m)
  movel([0.517428, -1.414134, -2.542415, -0.755840, 1.570796, 2.088224],accel_mss,speed_ms,0,blend_radius_m)
  movel([0.512611, -1.413625, -2.542799, -0.755965, 1.570796, 2.083408],accel_mss,speed_ms,0,blend_radius_m)
  movel([0.508038, -1.413190, -2.543127, -0.756071, 1.570796, 2.078835],accel_mss,speed_ms,0,blend_radius_m)
  movel([0.506156, -1.413233, -2.543095, -0.756061, 1.570796, 2.076952],accel_mss,speed_ms,0,blend_radius_m)
  movel([0.504193, -1.413515, -2.542883, -0.755992, 1.570796, 2.074989],accel_mss,speed_ms,0,blend_radius_m)
  movel([0.502203, -1.414101, -2.542440, -0.755849, 1.570796, 2.072999],accel_mss,speed_ms,0,blend_radius_m)
  movel([0.500246, -1.415056, -2.541717, -0.755616, 1.570796, 2.071042],accel_mss,speed_ms,0,blend_radius_m)
  movel([0.500537, -1.415781, -2.541168, -0.755441, 1.570796, 2.071333],accel_mss,speed_ms,0,blend_radius_m)
  movel([0.501483, -1.417705, -2.539705, -0.754979, 1.570796, 2.072279],accel_mss,speed_ms,0,blend_radius_m)
  movel([0.502598, -1.419225, -2.538546, -0.754618, 1.570796, 2.073394],accel_mss,speed_ms,0,blend_radius_m)
  movel([0.503882, -1.420340, -2.537694, -0.754355, 1.570796, 2.074679],accel_mss,speed_ms,0,blend_radius_m)
  movel([0.505338, -1.421051, -2.537149, -0.754189, 1.570796, 2.076135],accel_mss,speed_ms,0,blend_radius_m)
  movel([0.506925, -1.421402, -2.536880, -0.754107, 1.570796, 2.077721],accel_mss,speed_ms,0,blend_radius_m)
  movel([0.508596, -1.421433, -2.536856, -0.754100, 1.570796, 2.079392],accel_mss,speed_ms,0,blend_radius_m)
  movel([0.510358, -1.421144, -2.537077, -0.754167, 1.570796, 2.081154],accel_mss,speed_ms,0,blend_radius_m)
  movel([0.512210, -1.420535, -2.537544, -0.754310, 1.570796, 2.083007],accel_mss,speed_ms,0,blend_radius_m)
  movel([0.503399, -1.425618, -2.533634, -0.753138, 1.570796, 2.074195],accel_mss,speed_ms,0,blend_radius_m)
  movel([0.495562, -1.406301, -2.548292, -0.757796, 1.570796, 2.066359],accel_mss,speed_ms,0,blend_radius_m)
  movel([0.496458, -1.405765, -2.548690, -0.757933, 1.570796, 2.067255],accel_mss,speed_ms,0,blend_radius_m)
  speed_ms = 0.003
  movel([0.496458, -1.399421, -2.545759, -0.767209, 1.570796, 2.067255],accel_mss,speed_ms,0,blend_radius_m)
  speed_ms = 0.05
  movel([0.496458, -1.374956, -2.533748, -0.803685, 1.570796, 2.067255],accel_mss,speed_ms,0,blend_radius_m)
  #M_RunCode9
  movel([0.509832, -1.394517, -2.519590, -0.798282, 1.570796, 2.080628],accel_mss,speed_ms,0,blend_radius_m)
  #M_RunCode3
  movel([0.509832, -1.418608, -2.531358, -0.762423, 1.570796, 2.080628],accel_mss,speed_ms,0,blend_radius_m)
  speed_ms = 0.003
  movel([0.509832, -1.424848, -2.534228, -0.753313, 1.570796, 2.080628],accel_mss,speed_ms,0,blend_radius_m)
  speed_ms = 0.02
  movel([0.511489, -1.424174, -2.534748, -0.753467, 1.570796, 2.082285],accel_mss,speed_ms,0,blend_radius_m)
  movel([0.512932, -1.424174, -2.534749, -0.753467, 1.570796, 2.083728],accel_mss,speed_ms,0,blend_radius_m)
  movel([0.514055, -1.424738, -2.534313, -0.753338, 1.570796, 2.084852],accel_mss,speed_ms,0,blend_radius_m)
  movel([0.514744, -1.425759, -2.533524, -0.753105, 1.570796, 2.085541],accel_mss,speed_ms,0,blend_radius_m)
  movel([0.514937, -1.427058, -2.532519, -0.752812, 1.570796, 2.085734],accel_mss,speed_ms,0,blend_radius_m)
  movel([0.514570, -1.428467, -2.531425, -0.752498, 1.570796, 2.085366],accel_mss,speed_ms,0,blend_radius_m)
  movel([0.513651, -1.429811, -2.530378, -0.752200, 1.570796, 2.084447],accel_mss,speed_ms,0,blend_radius_m)
  movel([0.512178, -1.430921, -2.529512, -0.751956, 1.570796, 2.082975],accel_mss,speed_ms,0,blend_radius_m)
  movel([0.510814, -1.431527, -2.529039, -0.751824, 1.570796, 2.081610],accel_mss,speed_ms,0,blend_radius_m)
  movel([0.509686, -1.431709, -2.528896, -0.751784, 1.570796, 2.080483],accel_mss,speed_ms,0,blend_radius_m)
  movel([0.508526, -1.431985, -2.528680, -0.751724, 1.570796, 2.079322],accel_mss,speed_ms,0,blend_radius_m)
  movel([0.507878, -1.432525, -2.528258, -0.751607, 1.570796, 2.078675],accel_mss,speed_ms,0,blend_radius_m)
  movel([0.507463, -1.433272, -2.527672, -0.751446, 1.570796, 2.078259],accel_mss,speed_ms,0,blend_radius_m)
  movel([0.507312, -1.434096, -2.527024, -0.751269, 1.570796, 2.078108],accel_mss,speed_ms,0,blend_radius_m)
  movel([0.507458, -1.434872, -2.526414, -0.751103, 1.570796, 2.078254],accel_mss,speed_ms,0,blend_radius_m)
  movel([0.507953, -1.435723, -2.525744, -0.750922, 1.570796, 2.078749],accel_mss,speed_ms,0,blend_radius_m)
  movel([0.508675, -1.436345, -2.525253, -0.750791, 1.570796, 2.079471],accel_mss,speed_ms,0,blend_radius_m)
  movel([0.509623, -1.436739, -2.524942, -0.750708, 1.570796, 2.080419],accel_mss,speed_ms,0,blend_radius_m)
  movel([0.510802, -1.436903, -2.524813, -0.750674, 1.570796, 2.081598],accel_mss,speed_ms,0,blend_radius_m)
  movel([0.512138, -1.436832, -2.524869, -0.750689, 1.570796, 2.082934],accel_mss,speed_ms,0,blend_radius_m)
  movel([0.513565, -1.436513, -2.525120, -0.750756, 1.570796, 2.084362],accel_mss,speed_ms,0,blend_radius_m)
  movel([0.515084, -1.435949, -2.525565, -0.750874, 1.570796, 2.085880],accel_mss,speed_ms,0,blend_radius_m)
  movel([0.516698, -1.435139, -2.526204, -0.751046, 1.570796, 2.087494],accel_mss,speed_ms,0,blend_radius_m)
  movel([0.519231, -1.433363, -2.527600, -0.751426, 1.570796, 2.090027],accel_mss,speed_ms,0,blend_radius_m)
  movel([0.521287, -1.431158, -2.529327, -0.751904, 1.570796, 2.092083],accel_mss,speed_ms,0,blend_radius_m)
  movel([0.522111, -1.429901, -2.530308, -0.752180, 1.570796, 2.092907],accel_mss,speed_ms,0,blend_radius_m)
  movel([0.522761, -1.428555, -2.531356, -0.752478, 1.570796, 2.093557],accel_mss,speed_ms,0,blend_radius_m)
  movel([0.523550, -1.425589, -2.533656, -0.753144, 1.570796, 2.094347],accel_mss,speed_ms,0,blend_radius_m)
  movel([0.523563, -1.422338, -2.536162, -0.753890, 1.570796, 2.094359],accel_mss,speed_ms,0,blend_radius_m)
  movel([0.522702, -1.418890, -2.538801, -0.754697, 1.570796, 2.093498],accel_mss,speed_ms,0,blend_radius_m)
  movel([0.536409, -1.411195, -2.544631, -0.756564, 1.570796, 2.107206],accel_mss,speed_ms,0,blend_radius_m)
  movel([0.541481, -1.426097, -2.533263, -0.753029, 1.570796, 2.112277],accel_mss,speed_ms,0,blend_radius_m)
  movel([0.532657, -1.430934, -2.529502, -0.751953, 1.570796, 2.103453],accel_mss,speed_ms,0,blend_radius_m)
  movel([0.534565, -1.429219, -2.530840, -0.752331, 1.570796, 2.105361],accel_mss,speed_ms,0,blend_radius_m)
  movel([0.536127, -1.427136, -2.532458, -0.752795, 1.570796, 2.106923],accel_mss,speed_ms,0,blend_radius_m)
  movel([0.537258, -1.424789, -2.534274, -0.753326, 1.570796, 2.108054],accel_mss,speed_ms,0,blend_radius_m)
  movel([0.537883, -1.422280, -2.536206, -0.753903, 1.570796, 2.108679],accel_mss,speed_ms,0,blend_radius_m)
  movel([0.537943, -1.419703, -2.538181, -0.754505, 1.570796, 2.108740],accel_mss,speed_ms,0,blend_radius_m)
  movel([0.537390, -1.417164, -2.540116, -0.755108, 1.570796, 2.108186],accel_mss,speed_ms,0,blend_radius_m)
  movel([0.527316, -1.422769, -2.535830, -0.753790, 1.570796, 2.098112],accel_mss,speed_ms,0,blend_radius_m)
  movel([0.528081, -1.425831, -2.533469, -0.753089, 1.570796, 2.098877],accel_mss,speed_ms,0,blend_radius_m)
  movel([0.528248, -1.429067, -2.530958, -0.752364, 1.570796, 2.099044],accel_mss,speed_ms,0,blend_radius_m)
  movel([0.527721, -1.432302, -2.528432, -0.751655, 1.570796, 2.098517],accel_mss,speed_ms,0,blend_radius_m)
  movel([0.527164, -1.433857, -2.527212, -0.751320, 1.570796, 2.097961],accel_mss,speed_ms,0,blend_radius_m)
  movel([0.526409, -1.435373, -2.526019, -0.750996, 1.570796, 2.097205],accel_mss,speed_ms,0,blend_radius_m)
  movel([0.525443, -1.436802, -2.524892, -0.750695, 1.570796, 2.096240],accel_mss,speed_ms,0,blend_radius_m)
  movel([0.524250, -1.438100, -2.523865, -0.750423, 1.570796, 2.095047],accel_mss,speed_ms,0,blend_radius_m)
  movel([0.522831, -1.439271, -2.522937, -0.750181, 1.570796, 2.093627],accel_mss,speed_ms,0,blend_radius_m)
  movel([0.521184, -1.440313, -2.522109, -0.749967, 1.570796, 2.091980],accel_mss,speed_ms,0,blend_radius_m)
  movel([0.519462, -1.441152, -2.521441, -0.749796, 1.570796, 2.090259],accel_mss,speed_ms,0,blend_radius_m)
  movel([0.517815, -1.441718, -2.520990, -0.749681, 1.570796, 2.088611],accel_mss,speed_ms,0,blend_radius_m)
  movel([0.516241, -1.442010, -2.520758, -0.749622, 1.570796, 2.087037],accel_mss,speed_ms,0,blend_radius_m)
  movel([0.514737, -1.442027, -2.520744, -0.749618, 1.570796, 2.085533],accel_mss,speed_ms,0,blend_radius_m)
  movel([0.512027, -1.441410, -2.521235, -0.749743, 1.570796, 2.082823],accel_mss,speed_ms,0,blend_radius_m)
  movel([0.509772, -1.440037, -2.522328, -0.750023, 1.570796, 2.080568],accel_mss,speed_ms,0,blend_radius_m)
  movel([0.507999, -1.438092, -2.523871, -0.750425, 1.570796, 2.078795],accel_mss,speed_ms,0,blend_radius_m)
  movel([0.506745, -1.435763, -2.525712, -0.750914, 1.570796, 2.077541],accel_mss,speed_ms,0,blend_radius_m)
  movel([0.506251, -1.433952, -2.527137, -0.751299, 1.570796, 2.077048],accel_mss,speed_ms,0,blend_radius_m)
  movel([0.506099, -1.431918, -2.528732, -0.751738, 1.570796, 2.076896],accel_mss,speed_ms,0,blend_radius_m)
  movel([0.506342, -1.429826, -2.530367, -0.752196, 1.570796, 2.077139],accel_mss,speed_ms,0,blend_radius_m)
  movel([0.507041, -1.427845, -2.531908, -0.752636, 1.570796, 2.077837],accel_mss,speed_ms,0,blend_radius_m)
  movel([0.508200, -1.426135, -2.533234, -0.753020, 1.570796, 2.078996],accel_mss,speed_ms,0,blend_radius_m)
  movel([0.509832, -1.424848, -2.534228, -0.753313, 1.570796, 2.080628],accel_mss,speed_ms,0,blend_radius_m)
  speed_ms = 0.003
  movel([0.509832, -1.418608, -2.531358, -0.762423, 1.570796, 2.080628],accel_mss,speed_ms,0,blend_radius_m)
  speed_ms = 0.05
  movel([0.509832, -1.394517, -2.519590, -0.798282, 1.570796, 2.080628],accel_mss,speed_ms,0,blend_radius_m)
  #M_RunCode9
  movel([0.516305, -1.314337, -2.574318, -0.823734, 1.570796, 2.087102],accel_mss,speed_ms,0,blend_radius_m)
  #M_RunCode3
  movel([0.516305, -1.339873, -2.587103, -0.785413, 1.570796, 2.087102],accel_mss,speed_ms,0,blend_radius_m)
  speed_ms = 0.003
  movel([0.516305, -1.346521, -2.590228, -0.775640, 1.570796, 2.087102],accel_mss,speed_ms,0,blend_radius_m)
  speed_ms = 0.02
  movel([0.513548, -1.347042, -2.589884, -0.775463, 1.570796, 2.084344],accel_mss,speed_ms,0,blend_radius_m)
  movel([0.510875, -1.346999, -2.589913, -0.775478, 1.570796, 2.081671],accel_mss,speed_ms,0,blend_radius_m)
  movel([0.508340, -1.346491, -2.590247, -0.775650, 1.570796, 2.079137],accel_mss,speed_ms,0,blend_radius_m)
  movel([0.506001, -1.345611, -2.590828, -0.775951, 1.570796, 2.076797],accel_mss,speed_ms,0,blend_radius_m)
  movel([0.503917, -1.344448, -2.591592, -0.776349, 1.570796, 2.074714],accel_mss,speed_ms,0,blend_radius_m)
  movel([0.505499, -1.341258, -2.593679, -0.777451, 1.570796, 2.076296],accel_mss,speed_ms,0,blend_radius_m)
  movel([0.507990, -1.337853, -2.595893, -0.778644, 1.570796, 2.078787],accel_mss,speed_ms,0,blend_radius_m)
  movel([0.511138, -1.334531, -2.598036, -0.779822, 1.570796, 2.081935],accel_mss,speed_ms,0,blend_radius_m)
  movel([0.514668, -1.331614, -2.599906, -0.780869, 1.570796, 2.085464],accel_mss,speed_ms,0,blend_radius_m)
  movel([0.518306, -1.329423, -2.601303, -0.781663, 1.570796, 2.089103],accel_mss,speed_ms,0,blend_radius_m)
  movel([0.520076, -1.328700, -2.601763, -0.781926, 1.570796, 2.090873],accel_mss,speed_ms,0,blend_radius_m)
  movel([0.521766, -1.328278, -2.602031, -0.782080, 1.570796, 2.092562],accel_mss,speed_ms,0,blend_radius_m)
  movel([0.523340, -1.328199, -2.602081, -0.782109, 1.570796, 2.094136],accel_mss,speed_ms,0,blend_radius_m)
  movel([0.524763, -1.328501, -2.601889, -0.781999, 1.570796, 2.095559],accel_mss,speed_ms,0,blend_radius_m)
  movel([0.525997, -1.329219, -2.601433, -0.781737, 1.570796, 2.096794],accel_mss,speed_ms,0,blend_radius_m)
  movel([0.527006, -1.330396, -2.600683, -0.781309, 1.570796, 2.097802],accel_mss,speed_ms,0,blend_radius_m)
  movel([0.527760, -1.332639, -2.599250, -0.780500, 1.570796, 2.098556],accel_mss,speed_ms,0,blend_radius_m)
  movel([0.527519, -1.335157, -2.597633, -0.779599, 1.570796, 2.098315],accel_mss,speed_ms,0,blend_radius_m)
  movel([0.526404, -1.337846, -2.595897, -0.778646, 1.570796, 2.097200],accel_mss,speed_ms,0,blend_radius_m)
  movel([0.524533, -1.340601, -2.594108, -0.777680, 1.570796, 2.095329],accel_mss,speed_ms,0,blend_radius_m)
  movel([0.521851, -1.343405, -2.592276, -0.776708, 1.570796, 2.092647],accel_mss,speed_ms,0,blend_radius_m)
  movel([0.519091, -1.345342, -2.591004, -0.776043, 1.570796, 2.089887],accel_mss,speed_ms,0,blend_radius_m)
  movel([0.516305, -1.346521, -2.590228, -0.775640, 1.570796, 2.087102],accel_mss,speed_ms,0,blend_radius_m)
  speed_ms = 0.003
  movel([0.516305, -1.339873, -2.587103, -0.785413, 1.570796, 2.087102],accel_mss,speed_ms,0,blend_radius_m)
  speed_ms = 0.05
  movel([0.516305, -1.314337, -2.574318, -0.823734, 1.570796, 2.087102],accel_mss,speed_ms,0,blend_radius_m)
  #M_RunCode9
  movel([0.597942, -1.229032, -2.623495, -0.859862, 1.570796, 2.168738],accel_mss,speed_ms,0,blend_radius_m)
  #M_RunCode3
  movel([0.597942, -1.255774, -2.637397, -0.819217, 1.570796, 2.168738],accel_mss,speed_ms,0,blend_radius_m)
  speed_ms = 0.003
  movel([0.597942, -1.262779, -2.640805, -0.808805, 1.570796, 2.168738],accel_mss,speed_ms,0,blend_radius_m)
  speed_ms = 0.02
  movel([0.596894, -1.261660, -2.641421, -0.809308, 1.570796, 2.167691],accel_mss,speed_ms,0,blend_radius_m)
  movel([0.596292, -1.260135, -2.642257, -0.809997, 1.570796, 2.167089],accel_mss,speed_ms,0,blend_radius_m)
  movel([0.595945, -1.258401, -2.643204, -0.810784, 1.570796, 2.166742],accel_mss,speed_ms,0,blend_radius_m)
  movel([0.596749, -1.258183, -2.643323, -0.810883, 1.570796, 2.167545],accel_mss,speed_ms,0,blend_radius_m)
  movel([0.597204, -1.258524, -2.643137, -0.810728, 1.570796, 2.168000],accel_mss,speed_ms,0,blend_radius_m)
  movel([0.597776, -1.258868, -2.642950, -0.810571, 1.570796, 2.168573],accel_mss,speed_ms,0,blend_radius_m)
  movel([0.598925, -1.258663, -2.643062, -0.810665, 1.570796, 2.169721],accel_mss,speed_ms,0,blend_radius_m)
  movel([0.600214, -1.257940, -2.643455, -0.810993, 1.570796, 2.171010],accel_mss,speed_ms,0,blend_radius_m)
  movel([0.601457, -1.256991, -2.643972, -0.811426, 1.570796, 2.172254],accel_mss,speed_ms,0,blend_radius_m)
  movel([0.603161, -1.255619, -2.644717, -0.812053, 1.570796, 2.173957],accel_mss,speed_ms,0,blend_radius_m)
  movel([0.602874, -1.253352, -2.645942, -0.813094, 1.570796, 2.173670],accel_mss,speed_ms,0,blend_radius_m)
  movel([0.601964, -1.251870, -2.646741, -0.813779, 1.570796, 2.172760],accel_mss,speed_ms,0,blend_radius_m)
  movel([0.601218, -1.251531, -2.646923, -0.813935, 1.570796, 2.172014],accel_mss,speed_ms,0,blend_radius_m)
  movel([0.600247, -1.251523, -2.646927, -0.813939, 1.570796, 2.171044],accel_mss,speed_ms,0,blend_radius_m)
  movel([0.599029, -1.251890, -2.646730, -0.813769, 1.570796, 2.169825],accel_mss,speed_ms,0,blend_radius_m)
  movel([0.597542, -1.252677, -2.646306, -0.813406, 1.570796, 2.168338],accel_mss,speed_ms,0,blend_radius_m)
  movel([0.598140, -1.251122, -2.647142, -0.814125, 1.570796, 2.168937],accel_mss,speed_ms,0,blend_radius_m)
  movel([0.598832, -1.249785, -2.647858, -0.814745, 1.570796, 2.169629],accel_mss,speed_ms,0,blend_radius_m)
  movel([0.599250, -1.249313, -2.648111, -0.814965, 1.570796, 2.170047],accel_mss,speed_ms,0,blend_radius_m)
  movel([0.599737, -1.249037, -2.648258, -0.815094, 1.570796, 2.170533],accel_mss,speed_ms,0,blend_radius_m)
  movel([0.600972, -1.249250, -2.648145, -0.814994, 1.570796, 2.171768],accel_mss,speed_ms,0,blend_radius_m)
  movel([0.602804, -1.250721, -2.647357, -0.814311, 1.570796, 2.173600],accel_mss,speed_ms,0,blend_radius_m)
  movel([0.604041, -1.252805, -2.646238, -0.813347, 1.570796, 2.174838],accel_mss,speed_ms,0,blend_radius_m)
  movel([0.604296, -1.254029, -2.645577, -0.812783, 1.570796, 2.175092],accel_mss,speed_ms,0,blend_radius_m)
  movel([0.604226, -1.255355, -2.644860, -0.812174, 1.570796, 2.175022],accel_mss,speed_ms,0,blend_radius_m)
  movel([0.603781, -1.256760, -2.644098, -0.811531, 1.570796, 2.174577],accel_mss,speed_ms,0,blend_radius_m)
  movel([0.602901, -1.258228, -2.643299, -0.810862, 1.570796, 2.173697],accel_mss,speed_ms,0,blend_radius_m)
  movel([0.601698, -1.257363, -2.643770, -0.811256, 1.570796, 2.172494],accel_mss,speed_ms,0,blend_radius_m)
  movel([0.599628, -1.263287, -2.640525, -0.808577, 1.570796, 2.170424],accel_mss,speed_ms,0,blend_radius_m)
  movel([0.597942, -1.262779, -2.640805, -0.808805, 1.570796, 2.168738],accel_mss,speed_ms,0,blend_radius_m)
  speed_ms = 0.003
  movel([0.597942, -1.255774, -2.637397, -0.819217, 1.570796, 2.168738],accel_mss,speed_ms,0,blend_radius_m)
  speed_ms = 0.05
  movel([0.597942, -1.229032, -2.623495, -0.859862, 1.570796, 2.168738],accel_mss,speed_ms,0,blend_radius_m)
  #M_RunCode9
  movel([0.579642, -1.188227, -2.644020, -0.880142, 1.570796, 2.150438],accel_mss,speed_ms,0,blend_radius_m)
  #M_RunCode3
  movel([0.579642, -1.215387, -2.658461, -0.838541, 1.570796, 2.150438],accel_mss,speed_ms,0,blend_radius_m)
  speed_ms = 0.003
  movel([0.579642, -1.222524, -2.662006, -0.827859, 1.570796, 2.150438],accel_mss,speed_ms,0,blend_radius_m)
  speed_ms = 0.02
  movel([0.577022, -1.224440, -2.661039, -0.826909, 1.570796, 2.147818],accel_mss,speed_ms,0,blend_radius_m)
  movel([0.574289, -1.226131, -2.660183, -0.826075, 1.570796, 2.145085],accel_mss,speed_ms,0,blend_radius_m)
  movel([0.571472, -1.227559, -2.659458, -0.825372, 1.570796, 2.142268],accel_mss,speed_ms,0,blend_radius_m)
  movel([0.568597, -1.228697, -2.658878, -0.824814, 1.570796, 2.139394],accel_mss,speed_ms,0,blend_radius_m)
  movel([0.565700, -1.229516, -2.658460, -0.824413, 1.570796, 2.136497],accel_mss,speed_ms,0,blend_radius_m)
  movel([0.564244, -1.229631, -2.658401, -0.824357, 1.570796, 2.135041],accel_mss,speed_ms,0,blend_radius_m)
  movel([0.562805, -1.229508, -2.658464, -0.824417, 1.570796, 2.133601],accel_mss,speed_ms,0,blend_radius_m)
  movel([0.561504, -1.229410, -2.658514, -0.824465, 1.570796, 2.132300],accel_mss,speed_ms,0,blend_radius_m)
  movel([0.560481, -1.229587, -2.658423, -0.824379, 1.570796, 2.131277],accel_mss,speed_ms,0,blend_radius_m)
  movel([0.558726, -1.230798, -2.657803, -0.823787, 1.570796, 2.129523],accel_mss,speed_ms,0,blend_radius_m)
  movel([0.556412, -1.232758, -2.656796, -0.822835, 1.570796, 2.127209],accel_mss,speed_ms,0,blend_radius_m)
  movel([0.554012, -1.234828, -2.655728, -0.821833, 1.570796, 2.124808],accel_mss,speed_ms,0,blend_radius_m)
  movel([0.551985, -1.236376, -2.654926, -0.821087, 1.570796, 2.122782],accel_mss,speed_ms,0,blend_radius_m)
  movel([0.547977, -1.238644, -2.653745, -0.820000, 1.570796, 2.118773],accel_mss,speed_ms,0,blend_radius_m)
  movel([0.544398, -1.240097, -2.652986, -0.819306, 1.570796, 2.115194],accel_mss,speed_ms,0,blend_radius_m)
  movel([0.541206, -1.240817, -2.652608, -0.818963, 1.570796, 2.112002],accel_mss,speed_ms,0,blend_radius_m)
  movel([0.538365, -1.240879, -2.652576, -0.818934, 1.570796, 2.109162],accel_mss,speed_ms,0,blend_radius_m)
  movel([0.535843, -1.240360, -2.652848, -0.819181, 1.570796, 2.106640],accel_mss,speed_ms,0,blend_radius_m)
  movel([0.533609, -1.239331, -2.653386, -0.819671, 1.570796, 2.104405],accel_mss,speed_ms,0,blend_radius_m)
  movel([0.531632, -1.237863, -2.654152, -0.820373, 1.570796, 2.102428],accel_mss,speed_ms,0,blend_radius_m)
  movel([0.529879, -1.236029, -2.655106, -0.821254, 1.570796, 2.100675],accel_mss,speed_ms,0,blend_radius_m)
  movel([0.526938, -1.231549, -2.657418, -0.823422, 1.570796, 2.097735],accel_mss,speed_ms,0,blend_radius_m)
  movel([0.524569, -1.226471, -2.660011, -0.825907, 1.570796, 2.095365],accel_mss,speed_ms,0,blend_radius_m)
  movel([0.520659, -1.216918, -2.664808, -0.830663, 1.570796, 2.091456],accel_mss,speed_ms,0,blend_radius_m)
  movel([0.518428, -1.213081, -2.666706, -0.832602, 1.570796, 2.089224],accel_mss,speed_ms,0,blend_radius_m)
  movel([0.515335, -1.209045, -2.668685, -0.834659, 1.570796, 2.086131],accel_mss,speed_ms,0,blend_radius_m)
  movel([0.511503, -1.205059, -2.670621, -0.836709, 1.570796, 2.082299],accel_mss,speed_ms,0,blend_radius_m)
  movel([0.507065, -1.201369, -2.672397, -0.838622, 1.570796, 2.077861],accel_mss,speed_ms,0,blend_radius_m)
  movel([0.502159, -1.198230, -2.673897, -0.840262, 1.570796, 2.072956],accel_mss,speed_ms,0,blend_radius_m)
  movel([0.496940, -1.195882, -2.675012, -0.841496, 1.570796, 2.067736],accel_mss,speed_ms,0,blend_radius_m)
  movel([0.491568, -1.194564, -2.675634, -0.842190, 1.570796, 2.062364],accel_mss,speed_ms,0,blend_radius_m)
  movel([0.488877, -1.194367, -2.675727, -0.842295, 1.570796, 2.059673],accel_mss,speed_ms,0,blend_radius_m)
  movel([0.486213, -1.194509, -2.675660, -0.842220, 1.570796, 2.057010],accel_mss,speed_ms,0,blend_radius_m)
  movel([0.483345, -1.195020, -2.675419, -0.841950, 1.570796, 2.054141],accel_mss,speed_ms,0,blend_radius_m)
  movel([0.479904, -1.195948, -2.674980, -0.841461, 1.570796, 2.050700],accel_mss,speed_ms,0,blend_radius_m)
  movel([0.476084, -1.197324, -2.674328, -0.840737, 1.570796, 2.046881],accel_mss,speed_ms,0,blend_radius_m)
  movel([0.472083, -1.199167, -2.673450, -0.839771, 1.570796, 2.042879],accel_mss,speed_ms,0,blend_radius_m)
  movel([0.468106, -1.201491, -2.672339, -0.838559, 1.570796, 2.038903],accel_mss,speed_ms,0,blend_radius_m)
  movel([0.464346, -1.204310, -2.670983, -0.837096, 1.570796, 2.035143],accel_mss,speed_ms,0,blend_radius_m)
  movel([0.461005, -1.207635, -2.669371, -0.835382, 1.570796, 2.031801],accel_mss,speed_ms,0,blend_radius_m)
  movel([0.459551, -1.209487, -2.668469, -0.834433, 1.570796, 2.030347],accel_mss,speed_ms,0,blend_radius_m)
  movel([0.458275, -1.211469, -2.667499, -0.833421, 1.570796, 2.029072],accel_mss,speed_ms,0,blend_radius_m)
  movel([0.456868, -1.214575, -2.665969, -0.831845, 1.570796, 2.027664],accel_mss,speed_ms,0,blend_radius_m)
  movel([0.456436, -1.217215, -2.664661, -0.830513, 1.570796, 2.027232],accel_mss,speed_ms,0,blend_radius_m)
  movel([0.456869, -1.219435, -2.663554, -0.829400, 1.570796, 2.027665],accel_mss,speed_ms,0,blend_radius_m)
  movel([0.458058, -1.221279, -2.662631, -0.828479, 1.570796, 2.028855],accel_mss,speed_ms,0,blend_radius_m)
  movel([0.459898, -1.222788, -2.661873, -0.827728, 1.570796, 2.030695],accel_mss,speed_ms,0,blend_radius_m)
  movel([0.462283, -1.224006, -2.661259, -0.827124, 1.570796, 2.033080],accel_mss,speed_ms,0,blend_radius_m)
  movel([0.465113, -1.224973, -2.660770, -0.826646, 1.570796, 2.035910],accel_mss,speed_ms,0,blend_radius_m)
  movel([0.468284, -1.225732, -2.660385, -0.826271, 1.570796, 2.039080],accel_mss,speed_ms,0,blend_radius_m)
  movel([0.475240, -1.226770, -2.659859, -0.825760, 1.570796, 2.046037],accel_mss,speed_ms,0,blend_radius_m)
  movel([0.482357, -1.227408, -2.659534, -0.825446, 1.570796, 2.053153],accel_mss,speed_ms,0,blend_radius_m)
  movel([0.488838, -1.227905, -2.659282, -0.825202, 1.570796, 2.059634],accel_mss,speed_ms,0,blend_radius_m)
  movel([0.493890, -1.228508, -2.658974, -0.824907, 1.570796, 2.064686],accel_mss,speed_ms,0,blend_radius_m)
  movel([0.505738, -1.230607, -2.657901, -0.823881, 1.570796, 2.076534],accel_mss,speed_ms,0,blend_radius_m)
  movel([0.511921, -1.231970, -2.657202, -0.823217, 1.570796, 2.082717],accel_mss,speed_ms,0,blend_radius_m)
  movel([0.516504, -1.233414, -2.656458, -0.822517, 1.570796, 2.087301],accel_mss,speed_ms,0,blend_radius_m)
  movel([0.518076, -1.234279, -2.656012, -0.822098, 1.570796, 2.088872],accel_mss,speed_ms,0,blend_radius_m)
  movel([0.519386, -1.235379, -2.655443, -0.821567, 1.570796, 2.090182],accel_mss,speed_ms,0,blend_radius_m)
  movel([0.521257, -1.238203, -2.653975, -0.820211, 1.570796, 2.092053],accel_mss,speed_ms,0,blend_radius_m)
  movel([0.522204, -1.241706, -2.652142, -0.818541, 1.570796, 2.093000],accel_mss,speed_ms,0,blend_radius_m)
  movel([0.522330, -1.245700, -2.650034, -0.816655, 1.570796, 2.093126],accel_mss,speed_ms,0,blend_radius_m)
  movel([0.521719, -1.250008, -2.647739, -0.814642, 1.570796, 2.092515],accel_mss,speed_ms,0,blend_radius_m)
  movel([0.520464, -1.254463, -2.645343, -0.812583, 1.570796, 2.091261],accel_mss,speed_ms,0,blend_radius_m)
  movel([0.518657, -1.258899, -2.642933, -0.810557, 1.570796, 2.089453],accel_mss,speed_ms,0,blend_radius_m)
  movel([0.516384, -1.263149, -2.640601, -0.808638, 1.570796, 2.087180],accel_mss,speed_ms,0,blend_radius_m)
  movel([0.512966, -1.268127, -2.637843, -0.806419, 1.570796, 2.083763],accel_mss,speed_ms,0,blend_radius_m)
  movel([0.511285, -1.270089, -2.636747, -0.805553, 1.570796, 2.082081],accel_mss,speed_ms,0,blend_radius_m)
  movel([0.509602, -1.271748, -2.635817, -0.804824, 1.570796, 2.080398],accel_mss,speed_ms,0,blend_radius_m)
  movel([0.507914, -1.273139, -2.635034, -0.804216, 1.570796, 2.078710],accel_mss,speed_ms,0,blend_radius_m)
  movel([0.506206, -1.274294, -2.634383, -0.803712, 1.570796, 2.077003],accel_mss,speed_ms,0,blend_radius_m)
  movel([0.502694, -1.276047, -2.633391, -0.802951, 1.570796, 2.073491],accel_mss,speed_ms,0,blend_radius_m)
  movel([0.498988, -1.277272, -2.632695, -0.802422, 1.570796, 2.069785],accel_mss,speed_ms,0,blend_radius_m)
  movel([0.495015, -1.278237, -2.632146, -0.802006, 1.570796, 2.065811],accel_mss,speed_ms,0,blend_radius_m)
  movel([0.485989, -1.280424, -2.630897, -0.801068, 1.570796, 2.056786],accel_mss,speed_ms,0,blend_radius_m)
  movel([0.485520, -1.280580, -2.630807, -0.801001, 1.570796, 2.056316],accel_mss,speed_ms,0,blend_radius_m)
  movel([0.485666, -1.280674, -2.630754, -0.800961, 1.570796, 2.056462],accel_mss,speed_ms,0,blend_radius_m)
  movel([0.487481, -1.280709, -2.630734, -0.800946, 1.570796, 2.058278],accel_mss,speed_ms,0,blend_radius_m)
  movel([0.494960, -1.280418, -2.630900, -0.801070, 1.570796, 2.065757],accel_mss,speed_ms,0,blend_radius_m)
  movel([0.507345, -1.280018, -2.631129, -0.801242, 1.570796, 2.078141],accel_mss,speed_ms,0,blend_radius_m)
  movel([0.499978, -1.283403, -2.629186, -0.799800, 1.570796, 2.070774],accel_mss,speed_ms,0,blend_radius_m)
  movel([0.491789, -1.286806, -2.627217, -0.798365, 1.570796, 2.062585],accel_mss,speed_ms,0,blend_radius_m)
  movel([0.483076, -1.290163, -2.625261, -0.796964, 1.570796, 2.053873],accel_mss,speed_ms,0,blend_radius_m)
  movel([0.474132, -1.293395, -2.623365, -0.795629, 1.570796, 2.044928],accel_mss,speed_ms,0,blend_radius_m)
  movel([0.456695, -1.299180, -2.619936, -0.793272, 1.570796, 2.027491],accel_mss,speed_ms,0,blend_radius_m)
  movel([0.448774, -1.301552, -2.618518, -0.792319, 1.570796, 2.019570],accel_mss,speed_ms,0,blend_radius_m)
  movel([0.441757, -1.303456, -2.617375, -0.791558, 1.570796, 2.012554],accel_mss,speed_ms,0,blend_radius_m)
  movel([0.431851, -1.309800, -2.613530, -0.789059, 1.570796, 2.002647],accel_mss,speed_ms,0,blend_radius_m)
  movel([0.421831, -1.316724, -2.609274, -0.786391, 1.570796, 1.992627],accel_mss,speed_ms,0,blend_radius_m)
  movel([0.401801, -1.331301, -2.600106, -0.780982, 1.570796, 1.972598],accel_mss,speed_ms,0,blend_radius_m)
  movel([0.391928, -1.338485, -2.595483, -0.778421, 1.570796, 1.962724],accel_mss,speed_ms,0,blend_radius_m)
  movel([0.382219, -1.345307, -2.591028, -0.776055, 1.570796, 1.953015],accel_mss,speed_ms,0,blend_radius_m)
  movel([0.372717, -1.351560, -2.586887, -0.773941, 1.570796, 1.943514],accel_mss,speed_ms,0,blend_radius_m)
  movel([0.363451, -1.357045, -2.583212, -0.772132, 1.570796, 1.934247],accel_mss,speed_ms,0,blend_radius_m)
  movel([0.359862, -1.358887, -2.581968, -0.771534, 1.570796, 1.930658],accel_mss,speed_ms,0,blend_radius_m)
  movel([0.356459, -1.360365, -2.580966, -0.771058, 1.570796, 1.927255],accel_mss,speed_ms,0,blend_radius_m)
  movel([0.353262, -1.361481, -2.580208, -0.770700, 1.570796, 1.924058],accel_mss,speed_ms,0,blend_radius_m)
  movel([0.350287, -1.362242, -2.579690, -0.770457, 1.570796, 1.921083],accel_mss,speed_ms,0,blend_radius_m)
  movel([0.347552, -1.362646, -2.579414, -0.770328, 1.570796, 1.918348],accel_mss,speed_ms,0,blend_radius_m)
  movel([0.345075, -1.362696, -2.579381, -0.770312, 1.570796, 1.915871],accel_mss,speed_ms,0,blend_radius_m)
  movel([0.342872, -1.362394, -2.579587, -0.770408, 1.570796, 1.913669],accel_mss,speed_ms,0,blend_radius_m)
  movel([0.340968, -1.361741, -2.580031, -0.770617, 1.570796, 1.911764],accel_mss,speed_ms,0,blend_radius_m)
  movel([0.339380, -1.360734, -2.580716, -0.770939, 1.570796, 1.910176],accel_mss,speed_ms,0,blend_radius_m)
  movel([0.338129, -1.359371, -2.581640, -0.771378, 1.570796, 1.908925],accel_mss,speed_ms,0,blend_radius_m)
  movel([0.337240, -1.357654, -2.582801, -0.771934, 1.570796, 1.908036],accel_mss,speed_ms,0,blend_radius_m)
  movel([0.336731, -1.355578, -2.584199, -0.772612, 1.570796, 1.907527],accel_mss,speed_ms,0,blend_radius_m)
  movel([0.336630, -1.353141, -2.585833, -0.773416, 1.570796, 1.907426],accel_mss,speed_ms,0,blend_radius_m)
  movel([0.336961, -1.350336, -2.587702, -0.774351, 1.570796, 1.907758],accel_mss,speed_ms,0,blend_radius_m)
  movel([0.337751, -1.347162, -2.589805, -0.775422, 1.570796, 1.908547],accel_mss,speed_ms,0,blend_radius_m)
  movel([0.339028, -1.343612, -2.592141, -0.776637, 1.570796, 1.909824],accel_mss,speed_ms,0,blend_radius_m)
  movel([0.341742, -1.344682, -2.591438, -0.776269, 1.570796, 1.912538],accel_mss,speed_ms,0,blend_radius_m)
  movel([0.343130, -1.345114, -2.591154, -0.776121, 1.570796, 1.913927],accel_mss,speed_ms,0,blend_radius_m)
  movel([0.344676, -1.345158, -2.591125, -0.776106, 1.570796, 1.915472],accel_mss,speed_ms,0,blend_radius_m)
  movel([0.346035, -1.344767, -2.591383, -0.776240, 1.570796, 1.916831],accel_mss,speed_ms,0,blend_radius_m)
  movel([0.347734, -1.343954, -2.591916, -0.776519, 1.570796, 1.918530],accel_mss,speed_ms,0,blend_radius_m)
  movel([0.351976, -1.341266, -2.593674, -0.777449, 1.570796, 1.922772],accel_mss,speed_ms,0,blend_radius_m)
  movel([0.357043, -1.337507, -2.596116, -0.778766, 1.570796, 1.927840],accel_mss,speed_ms,0,blend_radius_m)
  movel([0.362567, -1.333082, -2.598966, -0.780340, 1.570796, 1.933364],accel_mss,speed_ms,0,blend_radius_m)
  movel([0.373437, -1.323927, -2.604779, -0.783683, 1.570796, 1.944233],accel_mss,speed_ms,0,blend_radius_m)
  movel([0.381366, -1.317245, -2.608951, -0.786193, 1.570796, 1.952162],accel_mss,speed_ms,0,blend_radius_m)
  movel([0.388476, -1.311890, -2.612252, -0.788247, 1.570796, 1.959272],accel_mss,speed_ms,0,blend_radius_m)
  movel([0.395654, -1.306512, -2.615530, -0.790348, 1.570796, 1.966450],accel_mss,speed_ms,0,blend_radius_m)
  movel([0.381370, -1.309251, -2.613865, -0.789273, 1.570796, 1.952166],accel_mss,speed_ms,0,blend_radius_m)
  movel([0.374008, -1.310378, -2.613177, -0.788834, 1.570796, 1.944804],accel_mss,speed_ms,0,blend_radius_m)
  movel([0.367029, -1.310844, -2.612893, -0.788653, 1.570796, 1.937825],accel_mss,speed_ms,0,blend_radius_m)
  movel([0.363806, -1.310705, -2.612977, -0.788706, 1.570796, 1.934602],accel_mss,speed_ms,0,blend_radius_m)
  movel([0.360824, -1.310256, -2.613252, -0.788881, 1.570796, 1.931621],accel_mss,speed_ms,0,blend_radius_m)
  movel([0.358134, -1.309443, -2.613748, -0.789198, 1.570796, 1.928931],accel_mss,speed_ms,0,blend_radius_m)
  movel([0.355783, -1.308218, -2.614494, -0.789677, 1.570796, 1.926580],accel_mss,speed_ms,0,blend_radius_m)
  movel([0.353822, -1.306527, -2.615520, -0.790342, 1.570796, 1.924618],accel_mss,speed_ms,0,blend_radius_m)
  movel([0.352299, -1.304316, -2.616857, -0.791216, 1.570796, 1.923095],accel_mss,speed_ms,0,blend_radius_m)
  movel([0.351269, -1.301526, -2.618534, -0.792329, 1.570796, 1.922065],accel_mss,speed_ms,0,blend_radius_m)
  movel([0.350788, -1.298100, -2.620580, -0.793709, 1.570796, 1.921584],accel_mss,speed_ms,0,blend_radius_m)
  movel([0.351065, -1.293682, -2.623196, -0.795511, 1.570796, 1.921861],accel_mss,speed_ms,0,blend_radius_m)
  movel([0.352267, -1.288871, -2.626016, -0.797502, 1.570796, 1.923064],accel_mss,speed_ms,0,blend_radius_m)
  movel([0.354317, -1.283816, -2.628948, -0.799625, 1.570796, 1.925114],accel_mss,speed_ms,0,blend_radius_m)
  movel([0.357137, -1.278675, -2.631896, -0.801818, 1.570796, 1.927933],accel_mss,speed_ms,0,blend_radius_m)
  movel([0.360638, -1.273617, -2.634765, -0.804007, 1.570796, 1.931434],accel_mss,speed_ms,0,blend_radius_m)
  movel([0.364731, -1.268811, -2.637461, -0.806117, 1.570796, 1.935527],accel_mss,speed_ms,0,blend_radius_m)
  movel([0.369319, -1.264437, -2.639891, -0.808062, 1.570796, 1.940116],accel_mss,speed_ms,0,blend_radius_m)
  movel([0.374298, -1.260683, -2.641957, -0.809749, 1.570796, 1.945094],accel_mss,speed_ms,0,blend_radius_m)
  movel([0.377131, -1.259236, -2.642749, -0.810404, 1.570796, 1.947928],accel_mss,speed_ms,0,blend_radius_m)
  movel([0.380273, -1.258241, -2.643292, -0.810856, 1.570796, 1.951069],accel_mss,speed_ms,0,blend_radius_m)
  movel([0.382709, -1.258072, -2.643384, -0.810933, 1.570796, 1.953505],accel_mss,speed_ms,0,blend_radius_m)
  movel([0.383349, -1.258412, -2.643199, -0.810779, 1.570796, 1.954145],accel_mss,speed_ms,0,blend_radius_m)
  movel([0.383433, -1.259095, -2.642825, -0.810468, 1.570796, 1.954230],accel_mss,speed_ms,0,blend_radius_m)
  movel([0.380956, -1.259840, -2.642419, -0.810131, 1.570796, 1.951753],accel_mss,speed_ms,0,blend_radius_m)
  movel([0.378830, -1.260730, -2.641931, -0.809728, 1.570796, 1.949626],accel_mss,speed_ms,0,blend_radius_m)
  movel([0.377041, -1.261742, -2.641376, -0.809271, 1.570796, 1.947837],accel_mss,speed_ms,0,blend_radius_m)
  movel([0.375579, -1.262851, -2.640765, -0.808772, 1.570796, 1.946376],accel_mss,speed_ms,0,blend_radius_m)
  movel([0.374434, -1.264036, -2.640112, -0.808241, 1.570796, 1.945230],accel_mss,speed_ms,0,blend_radius_m)
  movel([0.373598, -1.265267, -2.639431, -0.807690, 1.570796, 1.944394],accel_mss,speed_ms,0,blend_radius_m)
  movel([0.373055, -1.266527, -2.638733, -0.807129, 1.570796, 1.943852],accel_mss,speed_ms,0,blend_radius_m)
  movel([0.372794, -1.267793, -2.638029, -0.806567, 1.570796, 1.943590],accel_mss,speed_ms,0,blend_radius_m)
  movel([0.373071, -1.270249, -2.636657, -0.805482, 1.570796, 1.943867],accel_mss,speed_ms,0,blend_radius_m)
  movel([0.374329, -1.272465, -2.635414, -0.804510, 1.570796, 1.945125],accel_mss,speed_ms,0,blend_radius_m)
  movel([0.376477, -1.274273, -2.634395, -0.803721, 1.570796, 1.947274],accel_mss,speed_ms,0,blend_radius_m)
  movel([0.379421, -1.275509, -2.633696, -0.803184, 1.570796, 1.950217],accel_mss,speed_ms,0,blend_radius_m)
  movel([0.381486, -1.275833, -2.633512, -0.803044, 1.570796, 1.952283],accel_mss,speed_ms,0,blend_radius_m)
  movel([0.384144, -1.275893, -2.633478, -0.803018, 1.570796, 1.954940],accel_mss,speed_ms,0,blend_radius_m)
  movel([0.390929, -1.275336, -2.633794, -0.803260, 1.570796, 1.961725],accel_mss,speed_ms,0,blend_radius_m)
  movel([0.399145, -1.274093, -2.634497, -0.803800, 1.570796, 1.969941],accel_mss,speed_ms,0,blend_radius_m)
  movel([0.408170, -1.272397, -2.635452, -0.804540, 1.570796, 1.978967],accel_mss,speed_ms,0,blend_radius_m)
  movel([0.426138, -1.268530, -2.637618, -0.806241, 1.570796, 1.996934],accel_mss,speed_ms,0,blend_radius_m)
  movel([0.439778, -1.265327, -2.639398, -0.807664, 1.570796, 2.010574],accel_mss,speed_ms,0,blend_radius_m)
  movel([0.446653, -1.263702, -2.640296, -0.808390, 1.570796, 2.017449],accel_mss,speed_ms,0,blend_radius_m)
  movel([0.450380, -1.262704, -2.640847, -0.808839, 1.570796, 2.021177],accel_mss,speed_ms,0,blend_radius_m)
  movel([0.453248, -1.261690, -2.641404, -0.809295, 1.570796, 2.024044],accel_mss,speed_ms,0,blend_radius_m)
  movel([0.454045, -1.261244, -2.641649, -0.809496, 1.570796, 2.024841],accel_mss,speed_ms,0,blend_radius_m)
  movel([0.454380, -1.260839, -2.641871, -0.809679, 1.570796, 2.025176],accel_mss,speed_ms,0,blend_radius_m)
  movel([0.454045, -1.259931, -2.642368, -0.810089, 1.570796, 2.024842],accel_mss,speed_ms,0,blend_radius_m)
  movel([0.451999, -1.258087, -2.643375, -0.810926, 1.570796, 2.022795],accel_mss,speed_ms,0,blend_radius_m)
  movel([0.449347, -1.256735, -2.644111, -0.811543, 1.570796, 2.020143],accel_mss,speed_ms,0,blend_radius_m)
  movel([0.443372, -1.254172, -2.645500, -0.812717, 1.570796, 2.014168],accel_mss,speed_ms,0,blend_radius_m)
  movel([0.440612, -1.252287, -2.646516, -0.813586, 1.570796, 2.011408],accel_mss,speed_ms,0,blend_radius_m)
  movel([0.438385, -1.249535, -2.647992, -0.814862, 1.570796, 2.009181],accel_mss,speed_ms,0,blend_radius_m)
  movel([0.437562, -1.247720, -2.648961, -0.815708, 1.570796, 2.008358],accel_mss,speed_ms,0,blend_radius_m)
  movel([0.436977, -1.245555, -2.650111, -0.816723, 1.570796, 2.007773],accel_mss,speed_ms,0,blend_radius_m)
  movel([0.436670, -1.242989, -2.651467, -0.817933, 1.570796, 2.007466],accel_mss,speed_ms,0,blend_radius_m)
  movel([0.436681, -1.239971, -2.653052, -0.819366, 1.570796, 2.007477],accel_mss,speed_ms,0,blend_radius_m)
  movel([0.437316, -1.235744, -2.655254, -0.821392, 1.570796, 2.008112],accel_mss,speed_ms,0,blend_radius_m)
  movel([0.438687, -1.231516, -2.657435, -0.823438, 1.570796, 2.009483],accel_mss,speed_ms,0,blend_radius_m)
  movel([0.440716, -1.227296, -2.659592, -0.825501, 1.570796, 2.011512],accel_mss,speed_ms,0,blend_radius_m)
  movel([0.443317, -1.223105, -2.661713, -0.827571, 1.570796, 2.014113],accel_mss,speed_ms,0,blend_radius_m)
  movel([0.446402, -1.218956, -2.663794, -0.829640, 1.570796, 2.017198],accel_mss,speed_ms,0,blend_radius_m)
  movel([0.449879, -1.214871, -2.665823, -0.831695, 1.570796, 2.020676],accel_mss,speed_ms,0,blend_radius_m)
  movel([0.453661, -1.210866, -2.667794, -0.833729, 1.570796, 2.024457],accel_mss,speed_ms,0,blend_radius_m)
  movel([0.457648, -1.206965, -2.669697, -0.835727, 1.570796, 2.028444],accel_mss,speed_ms,0,blend_radius_m)
  movel([0.465502, -1.200094, -2.673008, -0.839287, 1.570796, 2.036298],accel_mss,speed_ms,0,blend_radius_m)
  movel([0.472694, -1.194722, -2.675560, -0.842107, 1.570796, 2.043490],accel_mss,speed_ms,0,blend_radius_m)
  movel([0.478876, -1.190772, -2.677416, -0.844201, 1.570796, 2.049672],accel_mss,speed_ms,0,blend_radius_m)
  movel([0.483706, -1.188154, -2.678638, -0.845597, 1.570796, 2.054502],accel_mss,speed_ms,0,blend_radius_m)
  movel([0.490842, -1.185110, -2.680048, -0.847231, 1.570796, 2.061638],accel_mss,speed_ms,0,blend_radius_m)
  movel([0.497686, -1.183106, -2.680972, -0.848312, 1.570796, 2.068482],accel_mss,speed_ms,0,blend_radius_m)
  movel([0.504156, -1.182124, -2.681422, -0.848843, 1.570796, 2.074952],accel_mss,speed_ms,0,blend_radius_m)
  movel([0.510164, -1.182133, -2.681418, -0.848838, 1.570796, 2.080960],accel_mss,speed_ms,0,blend_radius_m)
  movel([0.515631, -1.183101, -2.680974, -0.848314, 1.570796, 2.086427],accel_mss,speed_ms,0,blend_radius_m)
  movel([0.520488, -1.184983, -2.680107, -0.847299, 1.570796, 2.091284],accel_mss,speed_ms,0,blend_radius_m)
  movel([0.524665, -1.187729, -2.678835, -0.845825, 1.570796, 2.095461],accel_mss,speed_ms,0,blend_radius_m)
  movel([0.528098, -1.191289, -2.677174, -0.843925, 1.570796, 2.098894],accel_mss,speed_ms,0,blend_radius_m)
  movel([0.530502, -1.195143, -2.675361, -0.841885, 1.570796, 2.101298],accel_mss,speed_ms,0,blend_radius_m)
  movel([0.532446, -1.199330, -2.673373, -0.839687, 1.570796, 2.103242],accel_mss,speed_ms,0,blend_radius_m)
  movel([0.534273, -1.203503, -2.671372, -0.837514, 1.570796, 2.105069],accel_mss,speed_ms,0,blend_radius_m)
  movel([0.536326, -1.207327, -2.669521, -0.835541, 1.570796, 2.107122],accel_mss,speed_ms,0,blend_radius_m)
  movel([0.538939, -1.210481, -2.667983, -0.833925, 1.570796, 2.109736],accel_mss,speed_ms,0,blend_radius_m)
  movel([0.540562, -1.211705, -2.667383, -0.833301, 1.570796, 2.111358],accel_mss,speed_ms,0,blend_radius_m)
  movel([0.542447, -1.212646, -2.666920, -0.832823, 1.570796, 2.113243],accel_mss,speed_ms,0,blend_radius_m)
  movel([0.544640, -1.213263, -2.666616, -0.832509, 1.570796, 2.115437],accel_mss,speed_ms,0,blend_radius_m)
  movel([0.547183, -1.213519, -2.666491, -0.832380, 1.570796, 2.117979],accel_mss,speed_ms,0,blend_radius_m)
  movel([0.550121, -1.213374, -2.666562, -0.832453, 1.570796, 2.120918],accel_mss,speed_ms,0,blend_radius_m)
  movel([0.553499, -1.212787, -2.666851, -0.832751, 1.570796, 2.124295],accel_mss,speed_ms,0,blend_radius_m)
  movel([0.556579, -1.211810, -2.667331, -0.833247, 1.570796, 2.127376],accel_mss,speed_ms,0,blend_radius_m)
  movel([0.559294, -1.210416, -2.668015, -0.833958, 1.570796, 2.130090],accel_mss,speed_ms,0,blend_radius_m)
  movel([0.561634, -1.208684, -2.668861, -0.834844, 1.570796, 2.132430],accel_mss,speed_ms,0,blend_radius_m)
  movel([0.563602, -1.206696, -2.669828, -0.835865, 1.570796, 2.134398],accel_mss,speed_ms,0,blend_radius_m)
  movel([0.565188, -1.204534, -2.670875, -0.836981, 1.570796, 2.135984],accel_mss,speed_ms,0,blend_radius_m)
  movel([0.566381, -1.202285, -2.671958, -0.838146, 1.570796, 2.137177],accel_mss,speed_ms,0,blend_radius_m)
  movel([0.567177, -1.200036, -2.673036, -0.839318, 1.570796, 2.137974],accel_mss,speed_ms,0,blend_radius_m)
  movel([0.567566, -1.197874, -2.674066, -0.840449, 1.570796, 2.138363],accel_mss,speed_ms,0,blend_radius_m)
  movel([0.567537, -1.195891, -2.675007, -0.841491, 1.570796, 2.138334],accel_mss,speed_ms,0,blend_radius_m)
  movel([0.567081, -1.194180, -2.675816, -0.842393, 1.570796, 2.137877],accel_mss,speed_ms,0,blend_radius_m)
  movel([0.566186, -1.192833, -2.676450, -0.843106, 1.570796, 2.136982],accel_mss,speed_ms,0,blend_radius_m)
  movel([0.564844, -1.191944, -2.676867, -0.843577, 1.570796, 2.135641],accel_mss,speed_ms,0,blend_radius_m)
  movel([0.563052, -1.191600, -2.677028, -0.843760, 1.570796, 2.133849],accel_mss,speed_ms,0,blend_radius_m)
  movel([0.560804, -1.191900, -2.676888, -0.843601, 1.570796, 2.131600],accel_mss,speed_ms,0,blend_radius_m)
  movel([0.558093, -1.192931, -2.676404, -0.843054, 1.570796, 2.128890],accel_mss,speed_ms,0,blend_radius_m)
  movel([0.554924, -1.194773, -2.675536, -0.842080, 1.570796, 2.125721],accel_mss,speed_ms,0,blend_radius_m)
  movel([0.556610, -1.195119, -2.675373, -0.841898, 1.570796, 2.127406],accel_mss,speed_ms,0,blend_radius_m)
  movel([0.557788, -1.195805, -2.675048, -0.841536, 1.570796, 2.128585],accel_mss,speed_ms,0,blend_radius_m)
  movel([0.558453, -1.196777, -2.674587, -0.841025, 1.570796, 2.129249],accel_mss,speed_ms,0,blend_radius_m)
  movel([0.558600, -1.197985, -2.674013, -0.840390, 1.570796, 2.129397],accel_mss,speed_ms,0,blend_radius_m)
  movel([0.558222, -1.199381, -2.673348, -0.839660, 1.570796, 2.129018],accel_mss,speed_ms,0,blend_radius_m)
  movel([0.557315, -1.200912, -2.672616, -0.838861, 1.570796, 2.128111],accel_mss,speed_ms,0,blend_radius_m)
  movel([0.555876, -1.202526, -2.671842, -0.838021, 1.570796, 2.126673],accel_mss,speed_ms,0,blend_radius_m)
  movel([0.553898, -1.204176, -2.671047, -0.837166, 1.570796, 2.124695],accel_mss,speed_ms,0,blend_radius_m)
  movel([0.550290, -1.206402, -2.669970, -0.836016, 1.570796, 2.121086],accel_mss,speed_ms,0,blend_radius_m)
  movel([0.547035, -1.207591, -2.669393, -0.835405, 1.570796, 2.117832],accel_mss,speed_ms,0,blend_radius_m)
  movel([0.544145, -1.207851, -2.669267, -0.835272, 1.570796, 2.114941],accel_mss,speed_ms,0,blend_radius_m)
  movel([0.541645, -1.207282, -2.669543, -0.835564, 1.570796, 2.112441],accel_mss,speed_ms,0,blend_radius_m)
  movel([0.539557, -1.205976, -2.670177, -0.836236, 1.570796, 2.110353],accel_mss,speed_ms,0,blend_radius_m)
  movel([0.537910, -1.204027, -2.671119, -0.837243, 1.570796, 2.108706],accel_mss,speed_ms,0,blend_radius_m)
  movel([0.536737, -1.201525, -2.672323, -0.838541, 1.570796, 2.107533],accel_mss,speed_ms,0,blend_radius_m)
  movel([0.536065, -1.198563, -2.673738, -0.840088, 1.570796, 2.106861],accel_mss,speed_ms,0,blend_radius_m)
  movel([0.535937, -1.195223, -2.675323, -0.841843, 1.570796, 2.106734],accel_mss,speed_ms,0,blend_radius_m)
  movel([0.536381, -1.191604, -2.677027, -0.843758, 1.570796, 2.107178],accel_mss,speed_ms,0,blend_radius_m)
  movel([0.537442, -1.187791, -2.678806, -0.845792, 1.570796, 2.108239],accel_mss,speed_ms,0,blend_radius_m)
  movel([0.539152, -1.183888, -2.680612, -0.847889, 1.570796, 2.109948],accel_mss,speed_ms,0,blend_radius_m)
  movel([0.541552, -1.179986, -2.682401, -0.850003, 1.570796, 2.112349],accel_mss,speed_ms,0,blend_radius_m)
  movel([0.544677, -1.176190, -2.684125, -0.852074, 1.570796, 2.115473],accel_mss,speed_ms,0,blend_radius_m)
  movel([0.548563, -1.172611, -2.685737, -0.854041, 1.570796, 2.119359],accel_mss,speed_ms,0,blend_radius_m)
  movel([0.553237, -1.169359, -2.687190, -0.855840, 1.570796, 2.124033],accel_mss,speed_ms,0,blend_radius_m)
  movel([0.556716, -1.167424, -2.688050, -0.856915, 1.570796, 2.127512],accel_mss,speed_ms,0,blend_radius_m)
  movel([0.560175, -1.165805, -2.688766, -0.857818, 1.570796, 2.130971],accel_mss,speed_ms,0,blend_radius_m)
  movel([0.563582, -1.164501, -2.689341, -0.858547, 1.570796, 2.134378],accel_mss,speed_ms,0,blend_radius_m)
  movel([0.566909, -1.163527, -2.689769, -0.859093, 1.570796, 2.137705],accel_mss,speed_ms,0,blend_radius_m)
  movel([0.570124, -1.162882, -2.690052, -0.859455, 1.570796, 2.140920],accel_mss,speed_ms,0,blend_radius_m)
  movel([0.573200, -1.162575, -2.690187, -0.859628, 1.570796, 2.143996],accel_mss,speed_ms,0,blend_radius_m)
  movel([0.576107, -1.162609, -2.690172, -0.859608, 1.570796, 2.146904],accel_mss,speed_ms,0,blend_radius_m)
  movel([0.578818, -1.162983, -2.690008, -0.859398, 1.570796, 2.149615],accel_mss,speed_ms,0,blend_radius_m)
  movel([0.581302, -1.163704, -2.689691, -0.858994, 1.570796, 2.152098],accel_mss,speed_ms,0,blend_radius_m)
  movel([0.583535, -1.164767, -2.689223, -0.858398, 1.570796, 2.154331],accel_mss,speed_ms,0,blend_radius_m)
  movel([0.585487, -1.166179, -2.688601, -0.857609, 1.570796, 2.156283],accel_mss,speed_ms,0,blend_radius_m)
  movel([0.587135, -1.167937, -2.687823, -0.856630, 1.570796, 2.157931],accel_mss,speed_ms,0,blend_radius_m)
  movel([0.588451, -1.170036, -2.686889, -0.855464, 1.570796, 2.159247],accel_mss,speed_ms,0,blend_radius_m)
  movel([0.589417, -1.172474, -2.685798, -0.854116, 1.570796, 2.160213],accel_mss,speed_ms,0,blend_radius_m)
  movel([0.590003, -1.175252, -2.684549, -0.852588, 1.570796, 2.160799],accel_mss,speed_ms,0,blend_radius_m)
  movel([0.590189, -1.178365, -2.683139, -0.850885, 1.570796, 2.160985],accel_mss,speed_ms,0,blend_radius_m)
  movel([0.589574, -1.181811, -2.681566, -0.849012, 1.570796, 2.160371],accel_mss,speed_ms,0,blend_radius_m)
  movel([0.588252, -1.185738, -2.679758, -0.846893, 1.570796, 2.159048],accel_mss,speed_ms,0,blend_radius_m)
  movel([0.586944, -1.189146, -2.678176, -0.845067, 1.570796, 2.157740],accel_mss,speed_ms,0,blend_radius_m)
  movel([0.586359, -1.191054, -2.677285, -0.844051, 1.570796, 2.157155],accel_mss,speed_ms,0,blend_radius_m)
  movel([0.587040, -1.192001, -2.676840, -0.843547, 1.570796, 2.157837],accel_mss,speed_ms,0,blend_radius_m)
  movel([0.588600, -1.193122, -2.676314, -0.842953, 1.570796, 2.159397],accel_mss,speed_ms,0,blend_radius_m)
  movel([0.590319, -1.194358, -2.675732, -0.842299, 1.570796, 2.161116],accel_mss,speed_ms,0,blend_radius_m)
  movel([0.591488, -1.195637, -2.675127, -0.841624, 1.570796, 2.162284],accel_mss,speed_ms,0,blend_radius_m)
  movel([0.592342, -1.197884, -2.674061, -0.840443, 1.570796, 2.163138],accel_mss,speed_ms,0,blend_radius_m)
  movel([0.592701, -1.200280, -2.672919, -0.839190, 1.570796, 2.163498],accel_mss,speed_ms,0,blend_radius_m)
  movel([0.592600, -1.202789, -2.671715, -0.837884, 1.570796, 2.163396],accel_mss,speed_ms,0,blend_radius_m)
  movel([0.592076, -1.205371, -2.670470, -0.836548, 1.570796, 2.162873],accel_mss,speed_ms,0,blend_radius_m)
  movel([0.591168, -1.207992, -2.669198, -0.835199, 1.570796, 2.161965],accel_mss,speed_ms,0,blend_radius_m)
  movel([0.589913, -1.210611, -2.667919, -0.833859, 1.570796, 2.160709],accel_mss,speed_ms,0,blend_radius_m)
  movel([0.588347, -1.213196, -2.666649, -0.832543, 1.570796, 2.159143],accel_mss,speed_ms,0,blend_radius_m)
  movel([0.586503, -1.215712, -2.665407, -0.831270, 1.570796, 2.157299],accel_mss,speed_ms,0,blend_radius_m)
  movel([0.584414, -1.218129, -2.664206, -0.830054, 1.570796, 2.155210],accel_mss,speed_ms,0,blend_radius_m)
  movel([0.582117, -1.220409, -2.663067, -0.828913, 1.570796, 2.152913],accel_mss,speed_ms,0,blend_radius_m)
  movel([0.579642, -1.222524, -2.662006, -0.827859, 1.570796, 2.150438],accel_mss,speed_ms,0,blend_radius_m)
  speed_ms = 0.003
  movel([0.579642, -1.215387, -2.658461, -0.838541, 1.570796, 2.150438],accel_mss,speed_ms,0,blend_radius_m)
  speed_ms = 0.05
  movel([0.579642, -1.188227, -2.644020, -0.880142, 1.570796, 2.150438],accel_mss,speed_ms,0,blend_radius_m)
  #M_RunCode9
  movel([0.596137, -1.187267, -2.644481, -0.880641, 1.570796, 2.166934],accel_mss,speed_ms,0,blend_radius_m)
  #M_RunCode3
  movel([0.596137, -1.214436, -2.658934, -0.839019, 1.570796, 2.166934],accel_mss,speed_ms,0,blend_radius_m)
  speed_ms = 0.003
  movel([0.596137, -1.221575, -2.662482, -0.828331, 1.570796, 2.166934],accel_mss,speed_ms,0,blend_radius_m)
  speed_ms = 0.02
  movel([0.597154, -1.219391, -2.663576, -0.829422, 1.570796, 2.167950],accel_mss,speed_ms,0,blend_radius_m)
  movel([0.599787, -1.214948, -2.665785, -0.831656, 1.570796, 2.170584],accel_mss,speed_ms,0,blend_radius_m)
  movel([0.602168, -1.210593, -2.667928, -0.833868, 1.570796, 2.172964],accel_mss,speed_ms,0,blend_radius_m)
  movel([0.602865, -1.208522, -2.668940, -0.834927, 1.570796, 2.173661],accel_mss,speed_ms,0,blend_radius_m)
  movel([0.603016, -1.206558, -2.669895, -0.835936, 1.570796, 2.173812],accel_mss,speed_ms,0,blend_radius_m)
  movel([0.603407, -1.207742, -2.669319, -0.835327, 1.570796, 2.174204],accel_mss,speed_ms,0,blend_radius_m)
  movel([0.603576, -1.210185, -2.668128, -0.834076, 1.570796, 2.174373],accel_mss,speed_ms,0,blend_radius_m)
  movel([0.603088, -1.212680, -2.666903, -0.832805, 1.570796, 2.173884],accel_mss,speed_ms,0,blend_radius_m)
  movel([0.602148, -1.215212, -2.665654, -0.831522, 1.570796, 2.172944],accel_mss,speed_ms,0,blend_radius_m)
  movel([0.600959, -1.217766, -2.664387, -0.830236, 1.570796, 2.171755],accel_mss,speed_ms,0,blend_radius_m)
  movel([0.598640, -1.222881, -2.661826, -0.827682, 1.570796, 2.169437],accel_mss,speed_ms,0,blend_radius_m)
  movel([0.597906, -1.225418, -2.660545, -0.826426, 1.570796, 2.168702],accel_mss,speed_ms,0,blend_radius_m)
  movel([0.597718, -1.227918, -2.659275, -0.825196, 1.570796, 2.168514],accel_mss,speed_ms,0,blend_radius_m)
  movel([0.598102, -1.230478, -2.657967, -0.823943, 1.570796, 2.168898],accel_mss,speed_ms,0,blend_radius_m)
  movel([0.598455, -1.231764, -2.657307, -0.823317, 1.570796, 2.169252],accel_mss,speed_ms,0,blend_radius_m)
  movel([0.598870, -1.232373, -2.656994, -0.823021, 1.570796, 2.169666],accel_mss,speed_ms,0,blend_radius_m)
  movel([0.600319, -1.231856, -2.657260, -0.823273, 1.570796, 2.171116],accel_mss,speed_ms,0,blend_radius_m)
  movel([0.601499, -1.231491, -2.657448, -0.823450, 1.570796, 2.172295],accel_mss,speed_ms,0,blend_radius_m)
  movel([0.602659, -1.231352, -2.657519, -0.823518, 1.570796, 2.173455],accel_mss,speed_ms,0,blend_radius_m)
  movel([0.604714, -1.231628, -2.657377, -0.823383, 1.570796, 2.175510],accel_mss,speed_ms,0,blend_radius_m)
  movel([0.606050, -1.232208, -2.657079, -0.823102, 1.570796, 2.176846],accel_mss,speed_ms,0,blend_radius_m)
  movel([0.606821, -1.233046, -2.656648, -0.822695, 1.570796, 2.177617],accel_mss,speed_ms,0,blend_radius_m)
  movel([0.607181, -1.234106, -2.656101, -0.822182, 1.570796, 2.177978],accel_mss,speed_ms,0,blend_radius_m)
  movel([0.607287, -1.236739, -2.654737, -0.820913, 1.570796, 2.178084],accel_mss,speed_ms,0,blend_radius_m)
  movel([0.607597, -1.239812, -2.653135, -0.819442, 1.570796, 2.178393],accel_mss,speed_ms,0,blend_radius_m)
  movel([0.608795, -1.243509, -2.651193, -0.817687, 1.570796, 2.179591],accel_mss,speed_ms,0,blend_radius_m)
  movel([0.610154, -1.247071, -2.649306, -0.816012, 1.570796, 2.180950],accel_mss,speed_ms,0,blend_radius_m)
  movel([0.611286, -1.250750, -2.647342, -0.814297, 1.570796, 2.182082],accel_mss,speed_ms,0,blend_radius_m)
  movel([0.611821, -1.254783, -2.645170, -0.812436, 1.570796, 2.182617],accel_mss,speed_ms,0,blend_radius_m)
  movel([0.611711, -1.257149, -2.643886, -0.811353, 1.570796, 2.182507],accel_mss,speed_ms,0,blend_radius_m)
  movel([0.611315, -1.259601, -2.642549, -0.810239, 1.570796, 2.182111],accel_mss,speed_ms,0,blend_radius_m)
  movel([0.609958, -1.264636, -2.639781, -0.807972, 1.570796, 2.180754],accel_mss,speed_ms,0,blend_radius_m)
  movel([0.608326, -1.269652, -2.636992, -0.805745, 1.570796, 2.179122],accel_mss,speed_ms,0,blend_radius_m)
  movel([0.606990, -1.274409, -2.634318, -0.803662, 1.570796, 2.177786],accel_mss,speed_ms,0,blend_radius_m)
  movel([0.605753, -1.281997, -2.629995, -0.800397, 1.570796, 2.176549],accel_mss,speed_ms,0,blend_radius_m)
  movel([0.605318, -1.285203, -2.628146, -0.799039, 1.570796, 2.176115],accel_mss,speed_ms,0,blend_radius_m)
  movel([0.604698, -1.288274, -2.626364, -0.797751, 1.570796, 2.175494],accel_mss,speed_ms,0,blend_radius_m)
  movel([0.603676, -1.291397, -2.624539, -0.796453, 1.570796, 2.174472],accel_mss,speed_ms,0,blend_radius_m)
  movel([0.602027, -1.294756, -2.622562, -0.795071, 1.570796, 2.172823],accel_mss,speed_ms,0,blend_radius_m)
  movel([0.599536, -1.298533, -2.620322, -0.793534, 1.570796, 2.170332],accel_mss,speed_ms,0,blend_radius_m)
  movel([0.595996, -1.302903, -2.617707, -0.791779, 1.570796, 2.166793],accel_mss,speed_ms,0,blend_radius_m)
  movel([0.592835, -1.306280, -2.615670, -0.790439, 1.570796, 2.163631],accel_mss,speed_ms,0,blend_radius_m)
  movel([0.589695, -1.309180, -2.613909, -0.789301, 1.570796, 2.160491],accel_mss,speed_ms,0,blend_radius_m)
  movel([0.586579, -1.311629, -2.612412, -0.788348, 1.570796, 2.157375],accel_mss,speed_ms,0,blend_radius_m)
  movel([0.583483, -1.313660, -2.611165, -0.787564, 1.570796, 2.154280],accel_mss,speed_ms,0,blend_radius_m)
  movel([0.580417, -1.315300, -2.610155, -0.786934, 1.570796, 2.151213],accel_mss,speed_ms,0,blend_radius_m)
  movel([0.577377, -1.316574, -2.609367, -0.786448, 1.570796, 2.148173],accel_mss,speed_ms,0,blend_radius_m)
  movel([0.574370, -1.317506, -2.608789, -0.786093, 1.570796, 2.145167],accel_mss,speed_ms,0,blend_radius_m)
  movel([0.571398, -1.318122, -2.608407, -0.785860, 1.570796, 2.142194],accel_mss,speed_ms,0,blend_radius_m)
  movel([0.568468, -1.318443, -2.608207, -0.785738, 1.570796, 2.139264],accel_mss,speed_ms,0,blend_radius_m)
  movel([0.565579, -1.318496, -2.608175, -0.785718, 1.570796, 2.136375],accel_mss,speed_ms,0,blend_radius_m)
  movel([0.559951, -1.317876, -2.608560, -0.785953, 1.570796, 2.130747],accel_mss,speed_ms,0,blend_radius_m)
  movel([0.554561, -1.316436, -2.609453, -0.786501, 1.570796, 2.125357],accel_mss,speed_ms,0,blend_radius_m)
  movel([0.549456, -1.314345, -2.610744, -0.787301, 1.570796, 2.120252],accel_mss,speed_ms,0,blend_radius_m)
  movel([0.545034, -1.311851, -2.612276, -0.788262, 1.570796, 2.115830],accel_mss,speed_ms,0,blend_radius_m)
  movel([0.539445, -1.308537, -2.614300, -0.789552, 1.570796, 2.110242],accel_mss,speed_ms,0,blend_radius_m)
  movel([0.532912, -1.305260, -2.616287, -0.790842, 1.570796, 2.103708],accel_mss,speed_ms,0,blend_radius_m)
  movel([0.529370, -1.303898, -2.617109, -0.791382, 1.570796, 2.100166],accel_mss,speed_ms,0,blend_radius_m)
  movel([0.525685, -1.302862, -2.617732, -0.791795, 1.570796, 2.096481],accel_mss,speed_ms,0,blend_radius_m)
  movel([0.521902, -1.302260, -2.618094, -0.792035, 1.570796, 2.092698],accel_mss,speed_ms,0,blend_radius_m)
  movel([0.518055, -1.302190, -2.618136, -0.792063, 1.570796, 2.088851],accel_mss,speed_ms,0,blend_radius_m)
  movel([0.514187, -1.302756, -2.617796, -0.791837, 1.570796, 2.084983],accel_mss,speed_ms,0,blend_radius_m)
  movel([0.510347, -1.304052, -2.617016, -0.791321, 1.570796, 2.081143],accel_mss,speed_ms,0,blend_radius_m)
  movel([0.508448, -1.305004, -2.616442, -0.790944, 1.570796, 2.079244],accel_mss,speed_ms,0,blend_radius_m)
  movel([0.506574, -1.306175, -2.615734, -0.790481, 1.570796, 2.077370],accel_mss,speed_ms,0,blend_radius_m)
  movel([0.504730, -1.307571, -2.614887, -0.789931, 1.570796, 2.075526],accel_mss,speed_ms,0,blend_radius_m)
  movel([0.502921, -1.309207, -2.613892, -0.789290, 1.570796, 2.073718],accel_mss,speed_ms,0,blend_radius_m)
  movel([0.501155, -1.311093, -2.612741, -0.788556, 1.570796, 2.071951],accel_mss,speed_ms,0,blend_radius_m)
  movel([0.499434, -1.313236, -2.611426, -0.787727, 1.570796, 2.070231],accel_mss,speed_ms,0,blend_radius_m)
  movel([0.496162, -1.318337, -2.608274, -0.785778, 1.570796, 2.066959],accel_mss,speed_ms,0,blend_radius_m)
  movel([0.495202, -1.320841, -2.606714, -0.784835, 1.570796, 2.065999],accel_mss,speed_ms,0,blend_radius_m)
  movel([0.494709, -1.323337, -2.605150, -0.783902, 1.570796, 2.065505],accel_mss,speed_ms,0,blend_radius_m)
  movel([0.494716, -1.325803, -2.603598, -0.782989, 1.570796, 2.065512],accel_mss,speed_ms,0,blend_radius_m)
  movel([0.495255, -1.328208, -2.602075, -0.782106, 1.570796, 2.066052],accel_mss,speed_ms,0,blend_radius_m)
  movel([0.497997, -1.325115, -2.604031, -0.783242, 1.570796, 2.068793],accel_mss,speed_ms,0,blend_radius_m)
  movel([0.500907, -1.322290, -2.605807, -0.784292, 1.570796, 2.071703],accel_mss,speed_ms,0,blend_radius_m)
  movel([0.503955, -1.319744, -2.607398, -0.785247, 1.570796, 2.074751],accel_mss,speed_ms,0,blend_radius_m)
  movel([0.507111, -1.317490, -2.608799, -0.786100, 1.570796, 2.077907],accel_mss,speed_ms,0,blend_radius_m)
  movel([0.510338, -1.315540, -2.610007, -0.786843, 1.570796, 2.081134],accel_mss,speed_ms,0,blend_radius_m)
  movel([0.513610, -1.313904, -2.611015, -0.787470, 1.570796, 2.084407],accel_mss,speed_ms,0,blend_radius_m)
  movel([0.516892, -1.312597, -2.611819, -0.787973, 1.570796, 2.087688],accel_mss,speed_ms,0,blend_radius_m)
  movel([0.520150, -1.311628, -2.612413, -0.788348, 1.570796, 2.090947],accel_mss,speed_ms,0,blend_radius_m)
  movel([0.523355, -1.311006, -2.612794, -0.788590, 1.570796, 2.094151],accel_mss,speed_ms,0,blend_radius_m)
  movel([0.526466, -1.310742, -2.612955, -0.788692, 1.570796, 2.097263],accel_mss,speed_ms,0,blend_radius_m)
  movel([0.529460, -1.310840, -2.612895, -0.788654, 1.570796, 2.100256],accel_mss,speed_ms,0,blend_radius_m)
  movel([0.532300, -1.311310, -2.612608, -0.788472, 1.570796, 2.103097],accel_mss,speed_ms,0,blend_radius_m)
  movel([0.534953, -1.312159, -2.612087, -0.788143, 1.570796, 2.105749],accel_mss,speed_ms,0,blend_radius_m)
  movel([0.537390, -1.313392, -2.611330, -0.787667, 1.570796, 2.108186],accel_mss,speed_ms,0,blend_radius_m)
  movel([0.539582, -1.315011, -2.610333, -0.787045, 1.570796, 2.110379],accel_mss,speed_ms,0,blend_radius_m)
  movel([0.541497, -1.317017, -2.609093, -0.786279, 1.570796, 2.112294],accel_mss,speed_ms,0,blend_radius_m)
  movel([0.542800, -1.318916, -2.607914, -0.785559, 1.570796, 2.113596],accel_mss,speed_ms,0,blend_radius_m)
  movel([0.543796, -1.320943, -2.606650, -0.784796, 1.570796, 2.114592],accel_mss,speed_ms,0,blend_radius_m)
  movel([0.544494, -1.323084, -2.605309, -0.783996, 1.570796, 2.115290],accel_mss,speed_ms,0,blend_radius_m)
  movel([0.544913, -1.325319, -2.603903, -0.783167, 1.570796, 2.115709],accel_mss,speed_ms,0,blend_radius_m)
  movel([0.544973, -1.329999, -2.600936, -0.781453, 1.570796, 2.115769],accel_mss,speed_ms,0,blend_radius_m)
  movel([0.544083, -1.334844, -2.597835, -0.779710, 1.570796, 2.114879],accel_mss,speed_ms,0,blend_radius_m)
  movel([0.542361, -1.339725, -2.594678, -0.777986, 1.570796, 2.113157],accel_mss,speed_ms,0,blend_radius_m)
  movel([0.539915, -1.344510, -2.591551, -0.776328, 1.570796, 2.110711],accel_mss,speed_ms,0,blend_radius_m)
  movel([0.536845, -1.349085, -2.588532, -0.774771, 1.570796, 2.107641],accel_mss,speed_ms,0,blend_radius_m)
  movel([0.533259, -1.353330, -2.585706, -0.773353, 1.570796, 2.104055],accel_mss,speed_ms,0,blend_radius_m)
  movel([0.529245, -1.357135, -2.583151, -0.772103, 1.570796, 2.100041],accel_mss,speed_ms,0,blend_radius_m)
  movel([0.524898, -1.360391, -2.580949, -0.771049, 1.570796, 2.095694],accel_mss,speed_ms,0,blend_radius_m)
  movel([0.520303, -1.362992, -2.579179, -0.770218, 1.570796, 2.091099],accel_mss,speed_ms,0,blend_radius_m)
  movel([0.517936, -1.364013, -2.578482, -0.769895, 1.570796, 2.088733],accel_mss,speed_ms,0,blend_radius_m)
  movel([0.515539, -1.364832, -2.577921, -0.769636, 1.570796, 2.086335],accel_mss,speed_ms,0,blend_radius_m)
  movel([0.513120, -1.365430, -2.577511, -0.769448, 1.570796, 2.083916],accel_mss,speed_ms,0,blend_radius_m)
  movel([0.510687, -1.365799, -2.577258, -0.769332, 1.570796, 2.081483],accel_mss,speed_ms,0,blend_radius_m)
  movel([0.508250, -1.365922, -2.577173, -0.769293, 1.570796, 2.079046],accel_mss,speed_ms,0,blend_radius_m)
  movel([0.505818, -1.365788, -2.577266, -0.769335, 1.570796, 2.076614],accel_mss,speed_ms,0,blend_radius_m)
  movel([0.503402, -1.365377, -2.577547, -0.769464, 1.570796, 2.074198],accel_mss,speed_ms,0,blend_radius_m)
  movel([0.501009, -1.364680, -2.578025, -0.769684, 1.570796, 2.071806],accel_mss,speed_ms,0,blend_radius_m)
  movel([0.498647, -1.363680, -2.578709, -0.770000, 1.570796, 2.069443],accel_mss,speed_ms,0,blend_radius_m)
  movel([0.496327, -1.362360, -2.579610, -0.770419, 1.570796, 2.067123],accel_mss,speed_ms,0,blend_radius_m)
  movel([0.494743, -1.360953, -2.580567, -0.770869, 1.570796, 2.065539],accel_mss,speed_ms,0,blend_radius_m)
  movel([0.490867, -1.356572, -2.583531, -0.772287, 1.570796, 2.061664],accel_mss,speed_ms,0,blend_radius_m)
  movel([0.488474, -1.353182, -2.585805, -0.773402, 1.570796, 2.059270],accel_mss,speed_ms,0,blend_radius_m)
  movel([0.485996, -1.348940, -2.588629, -0.774820, 1.570796, 2.056792],accel_mss,speed_ms,0,blend_radius_m)
  movel([0.483593, -1.343799, -2.592018, -0.776572, 1.570796, 2.054390],accel_mss,speed_ms,0,blend_radius_m)
  movel([0.481444, -1.337704, -2.595989, -0.778696, 1.570796, 2.052240],accel_mss,speed_ms,0,blend_radius_m)
  movel([0.480362, -1.333157, -2.598918, -0.780314, 1.570796, 2.051158],accel_mss,speed_ms,0,blend_radius_m)
  movel([0.479844, -1.328776, -2.601714, -0.781898, 1.570796, 2.050640],accel_mss,speed_ms,0,blend_radius_m)
  movel([0.479827, -1.324575, -2.604371, -0.783442, 1.570796, 2.050623],accel_mss,speed_ms,0,blend_radius_m)
  movel([0.480249, -1.320573, -2.606881, -0.784935, 1.570796, 2.051046],accel_mss,speed_ms,0,blend_radius_m)
  movel([0.481050, -1.316778, -2.609241, -0.786370, 1.570796, 2.051846],accel_mss,speed_ms,0,blend_radius_m)
  movel([0.482155, -1.313216, -2.611439, -0.787735, 1.570796, 2.052951],accel_mss,speed_ms,0,blend_radius_m)
  movel([0.483501, -1.309902, -2.613468, -0.789019, 1.570796, 2.054298],accel_mss,speed_ms,0,blend_radius_m)
  movel([0.485016, -1.306856, -2.615321, -0.790212, 1.570796, 2.055813],accel_mss,speed_ms,0,blend_radius_m)
  movel([0.488266, -1.301650, -2.618460, -0.792279, 1.570796, 2.059062],accel_mss,speed_ms,0,blend_radius_m)
